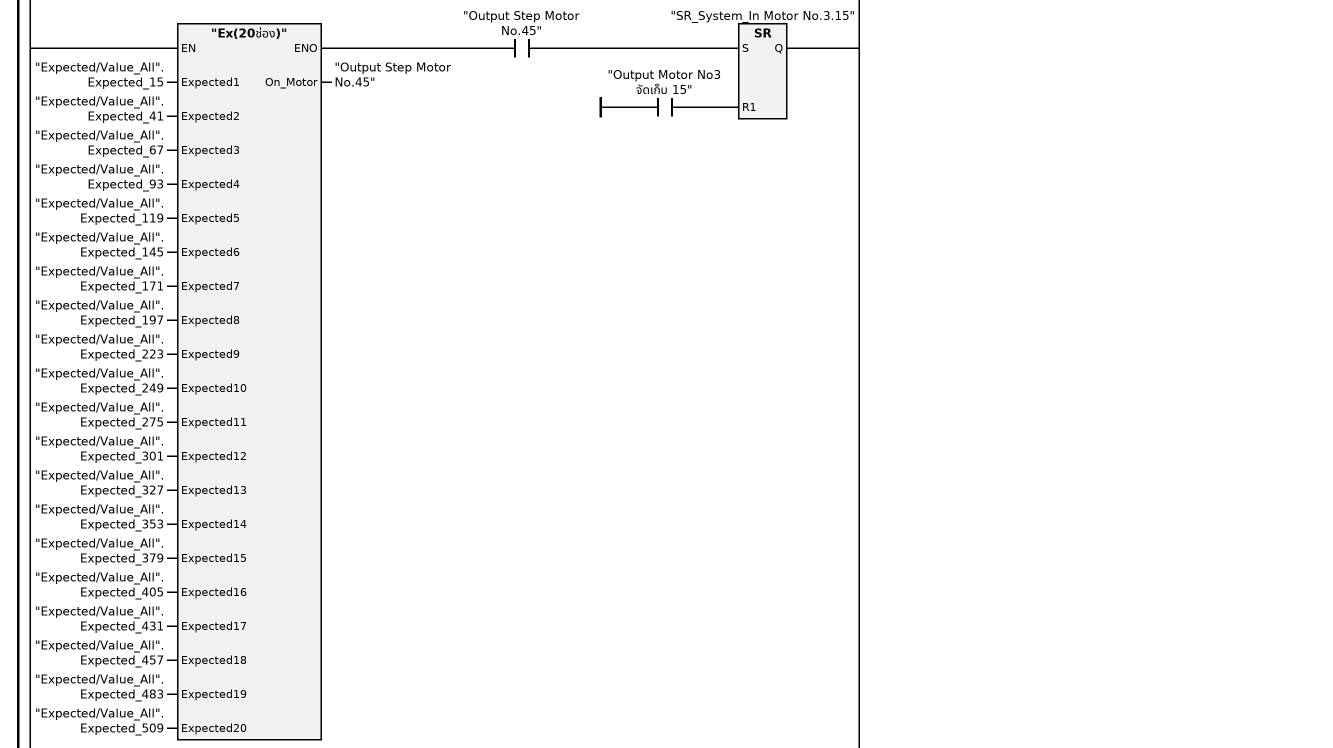
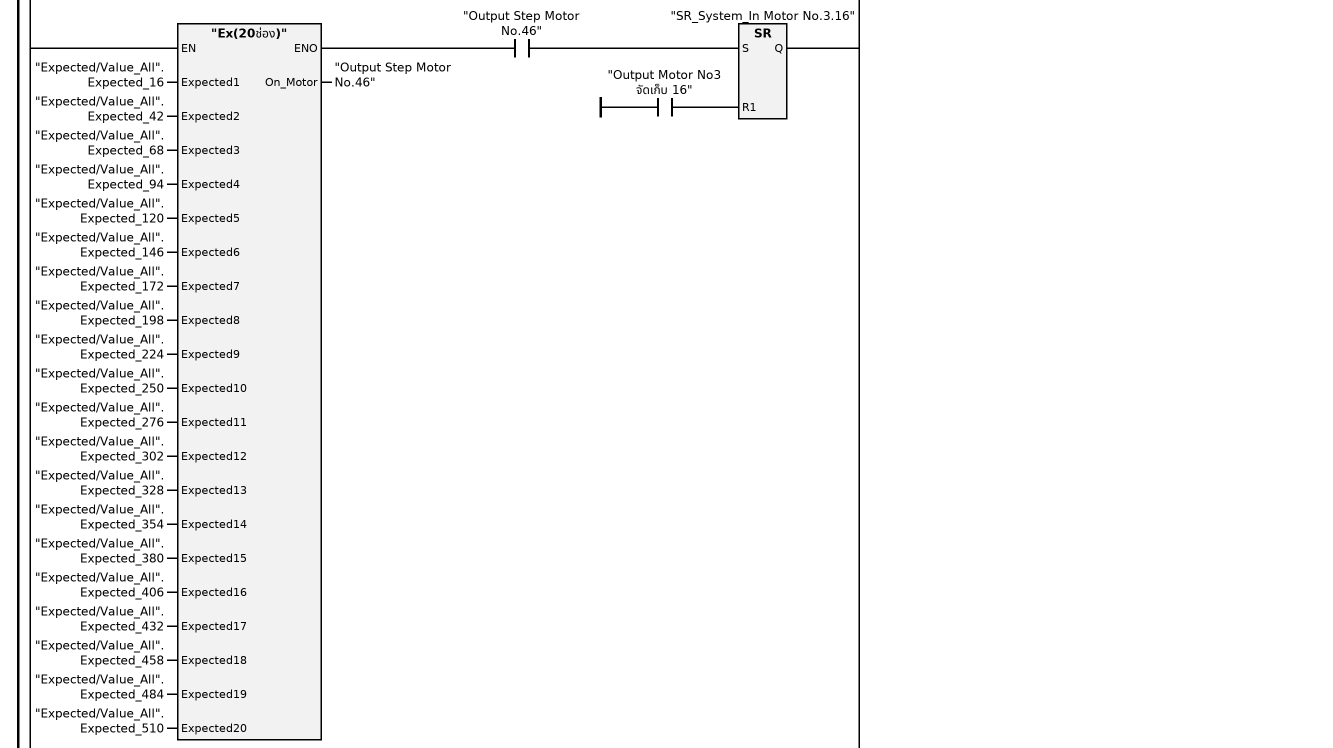
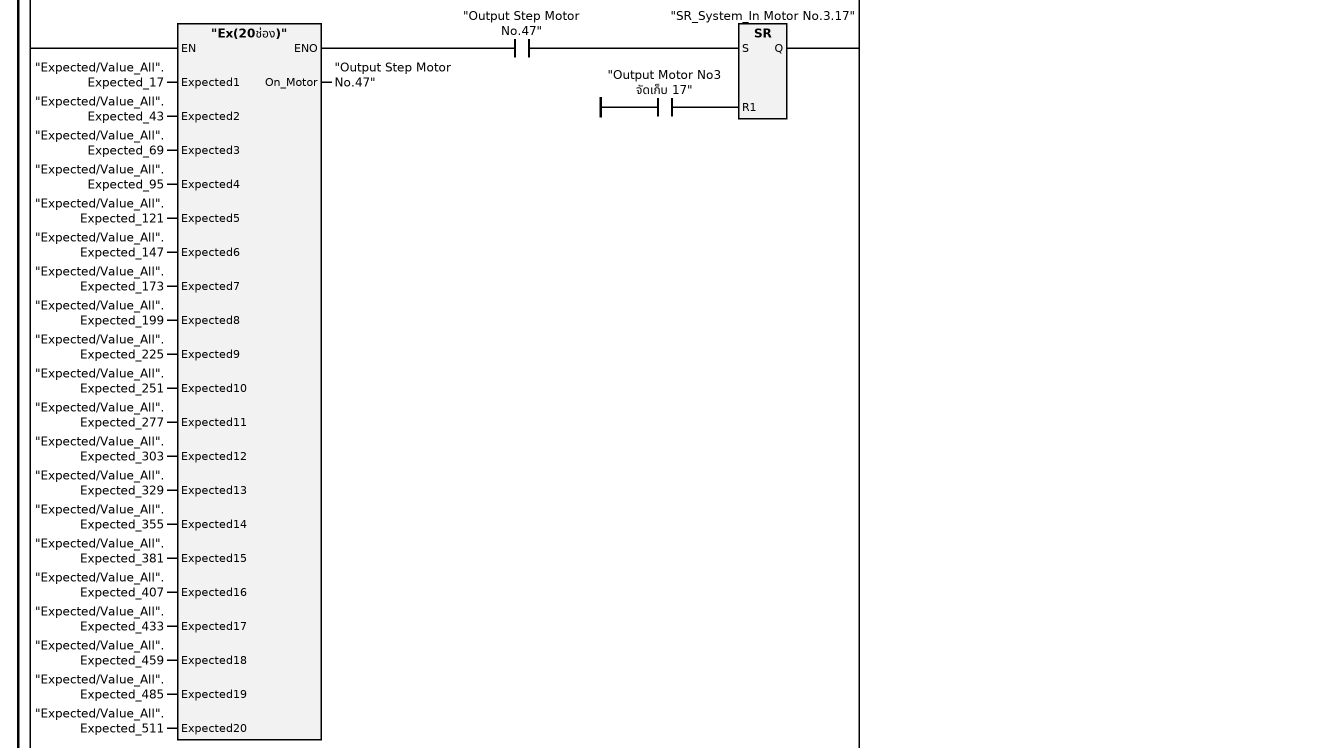
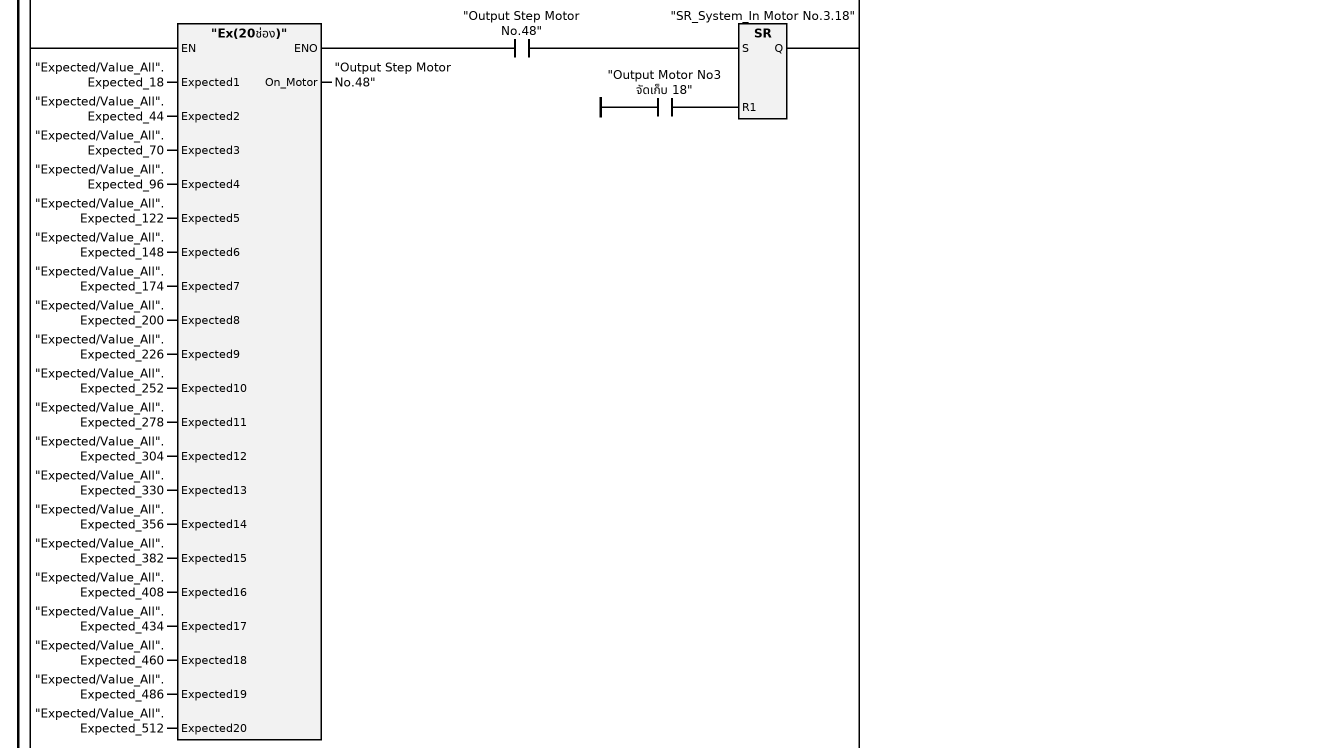
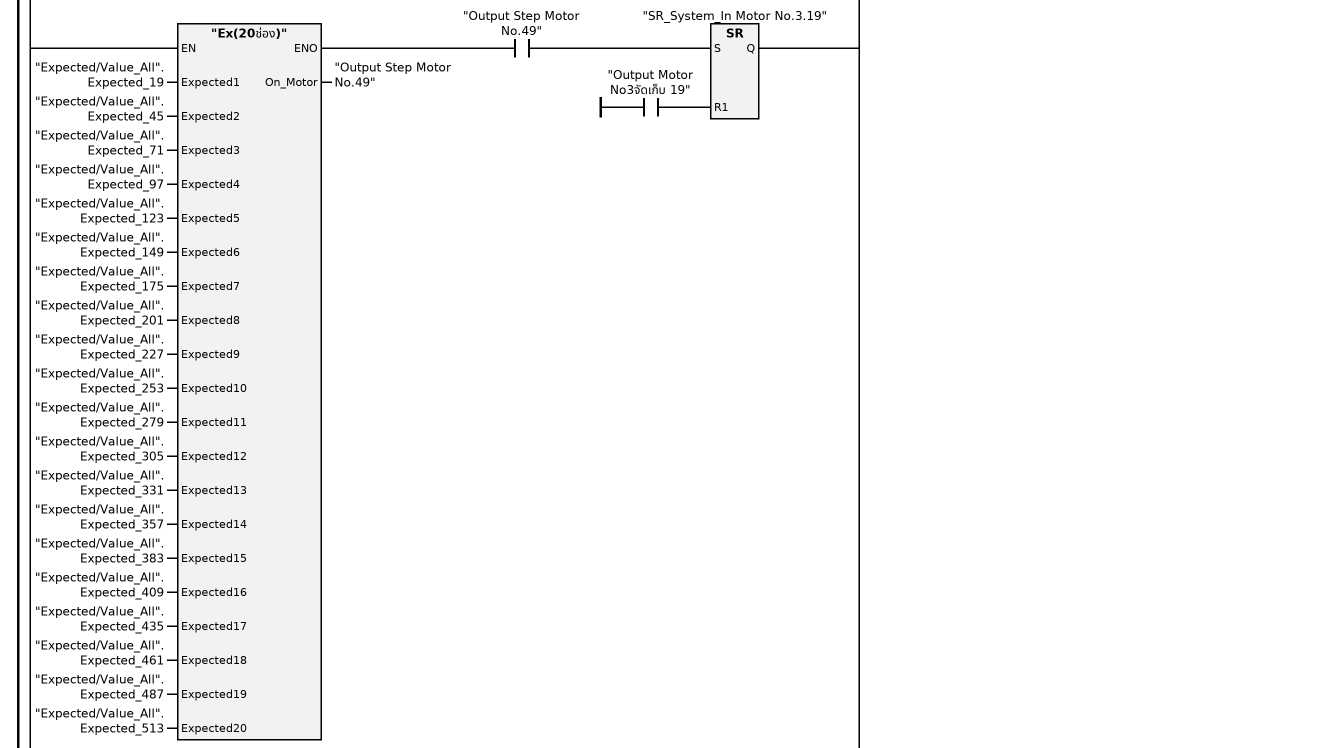
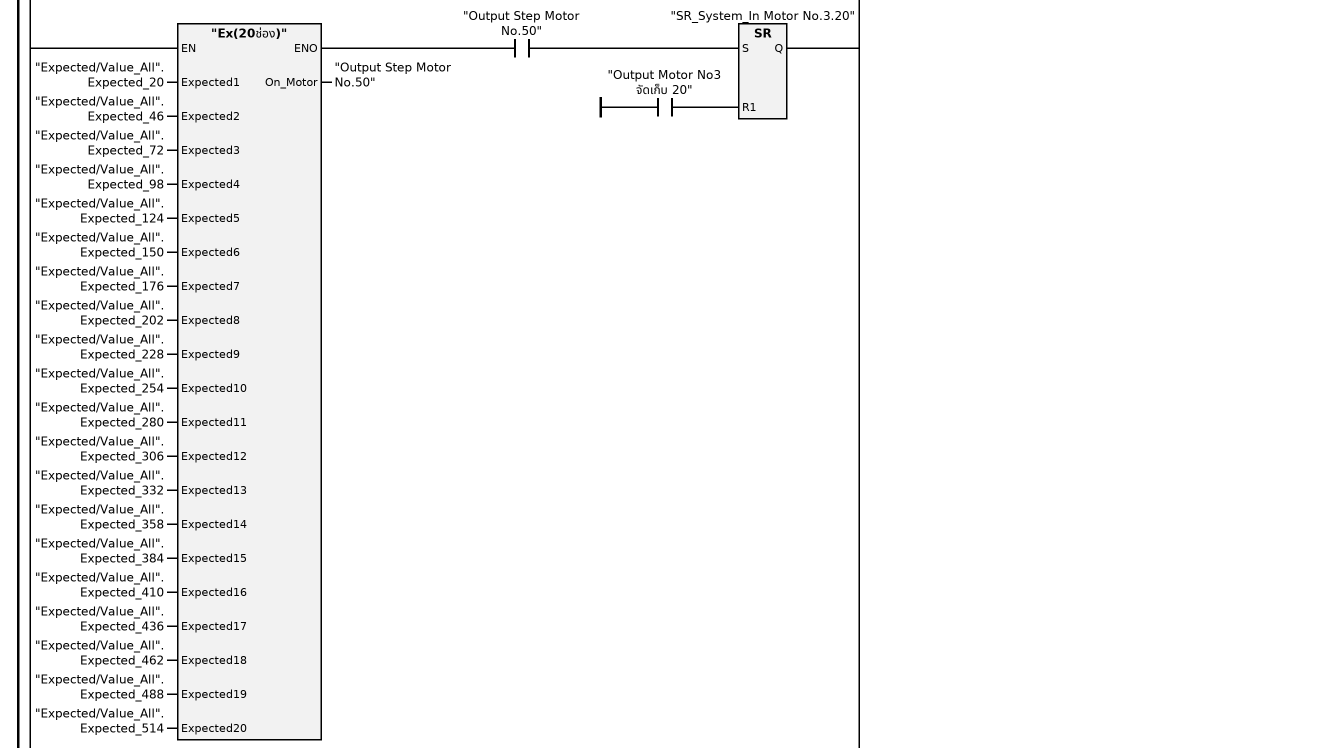
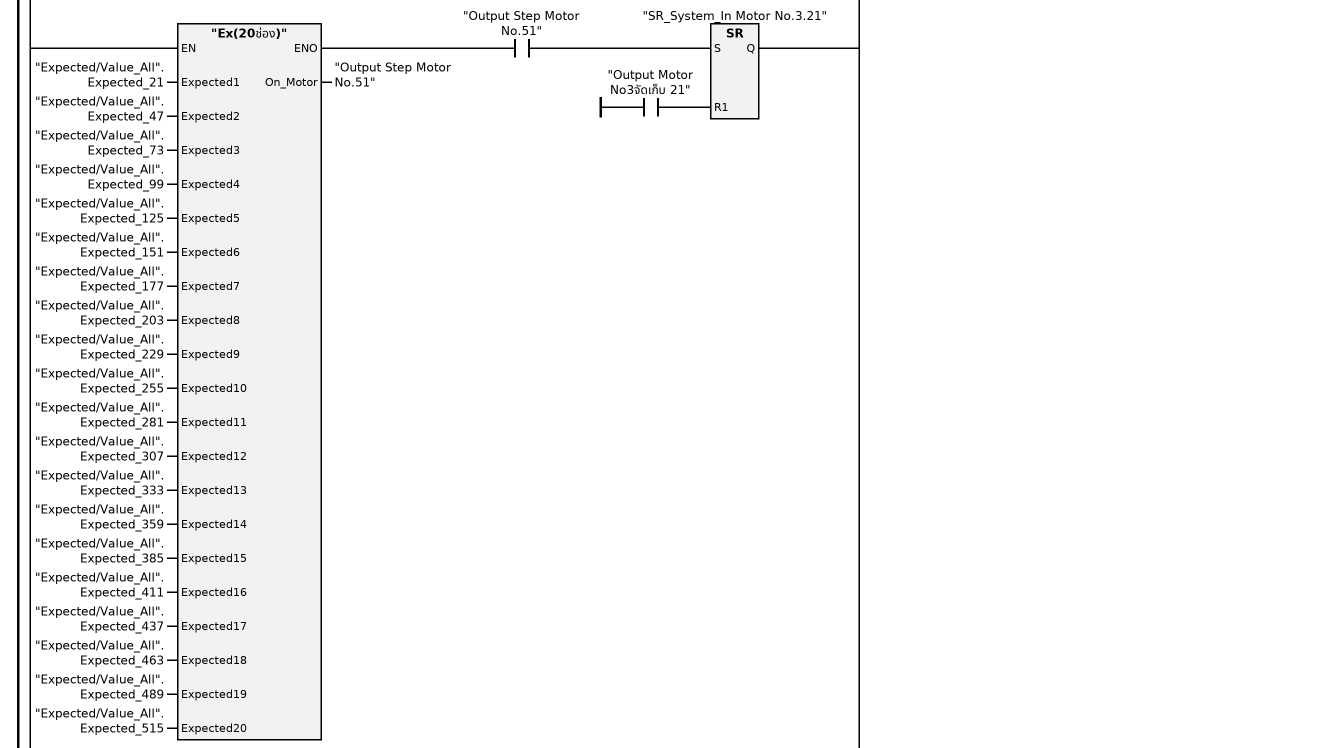
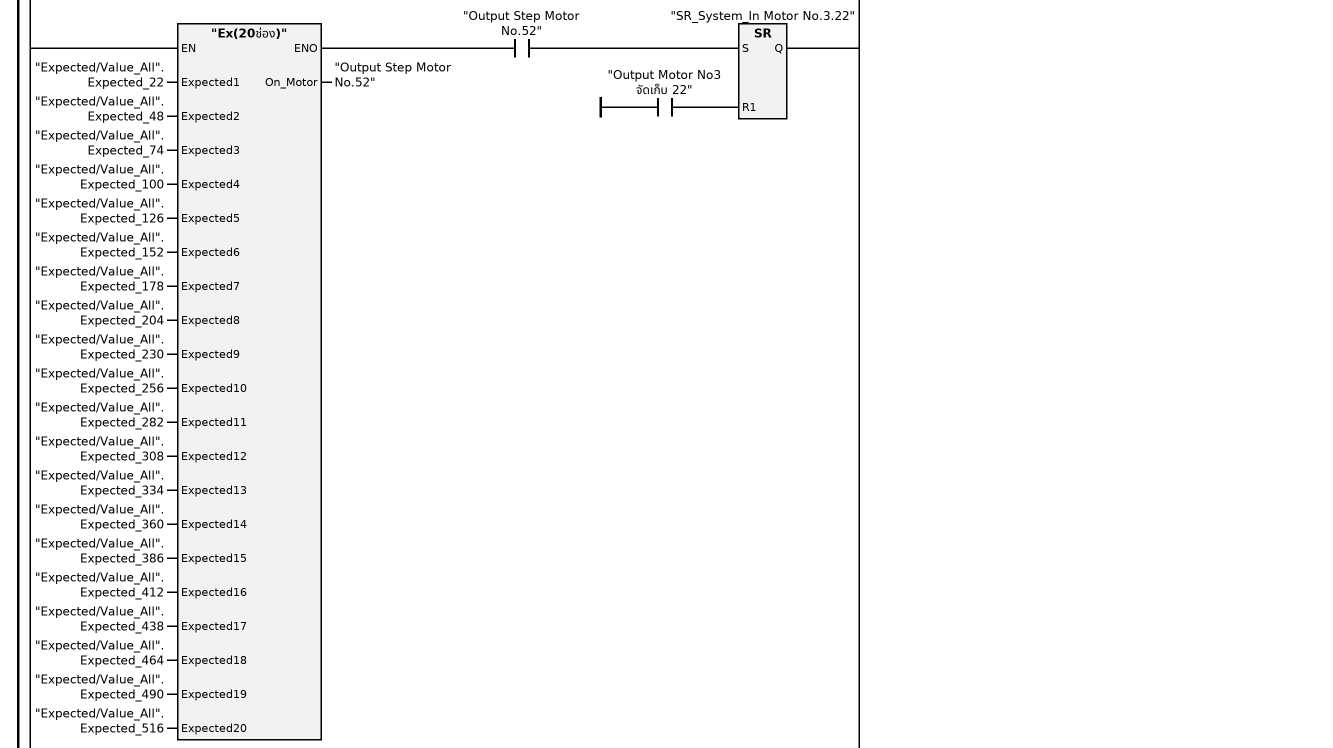
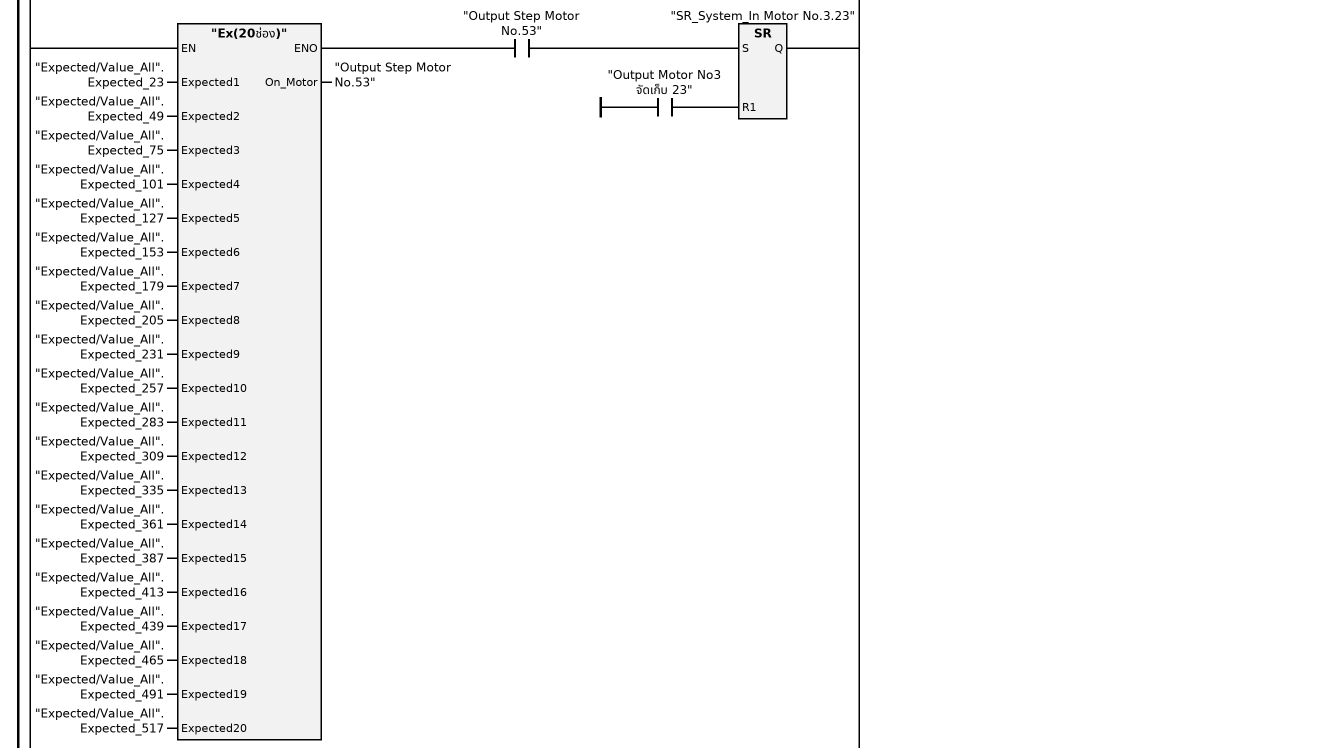
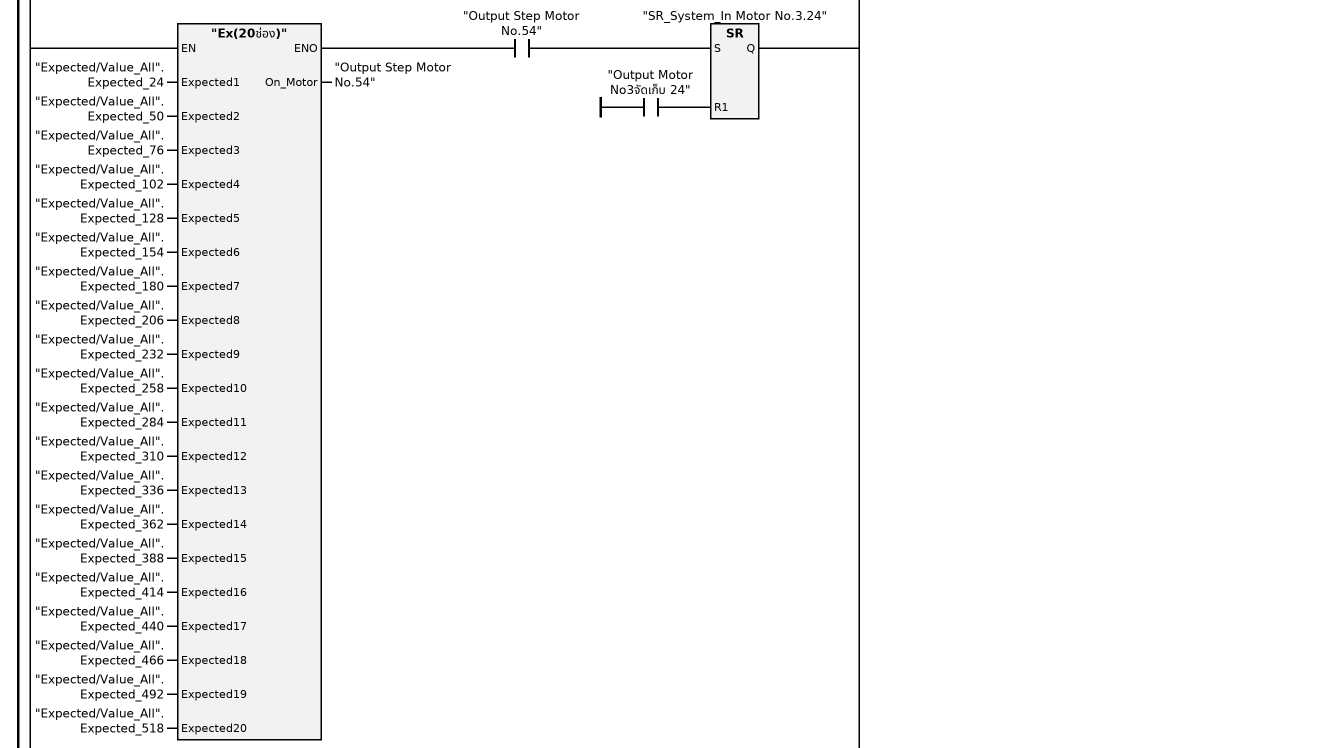
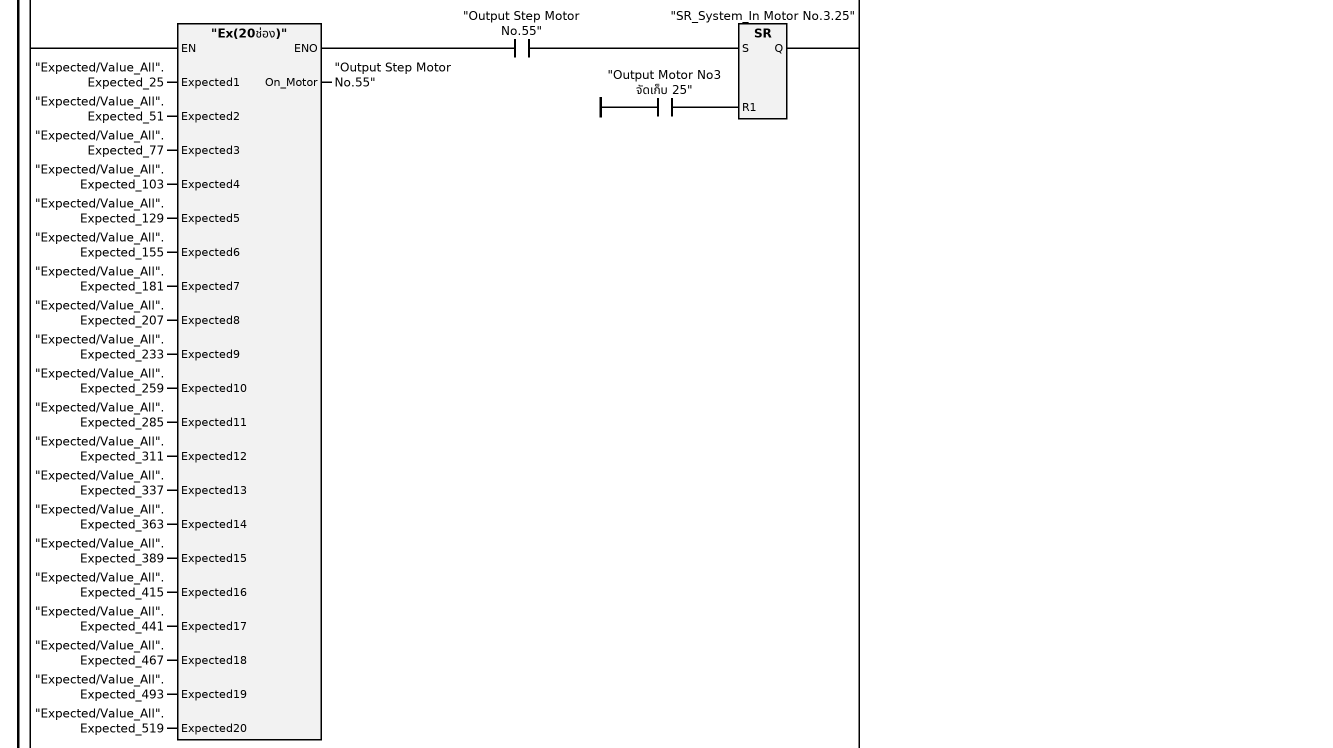
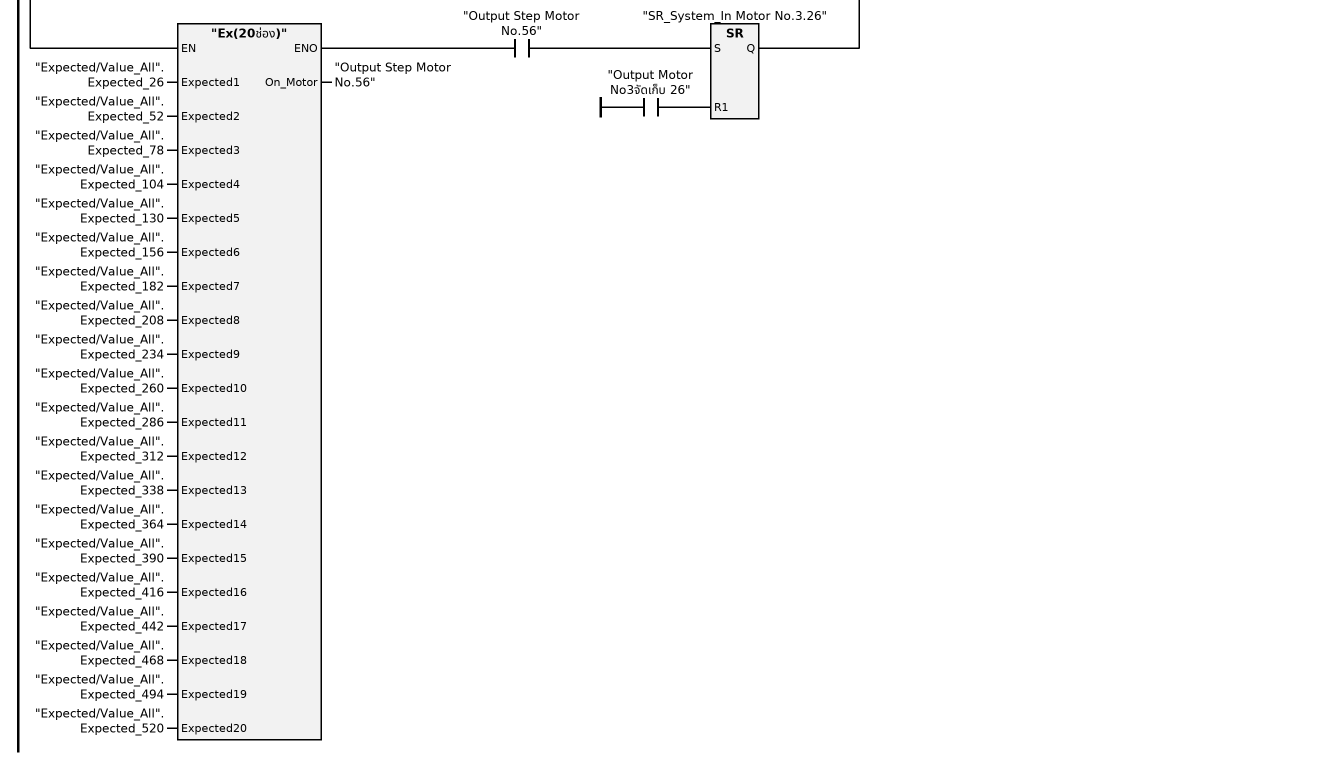
   "Ex(20ช่อง)"(Expected1 := "Expected/Value_All".Expected_1,
                Expected2 := "Expected/Value_All".Expected_27,
                Expected3 := "Expected/Value_All".Expected_53,
                Expected4 := "Expected/Value_All".Expected_79,
                Expected5 := "Expected/Value_All".Expected_105,
                Expected6 := "Expected/Value_All".Expected_131,
                Expected7 := "Expected/Value_All".Expected_157,
                Expected8 := "Expected/Value_All".Expected_183,
                Expected9 := "Expected/Value_All".Expected_209,
                Expected10 := "Expected/Value_All".Expected_235,
                Expected11 := "Expected/Value_All".Expected_261,
                Expected12 := "Expected/Value_All".Expected_287,
                Expected13 := "Expected/Value_All".Expected_313,
                Expected14 := "Expected/Value_All".Expected_339,
                Expected15 := "Expected/Value_All".Expected_365,
                Expected16 := "Expected/Value_All".Expected_391,
                Expected17 := "Expected/Value_All".Expected_417,
                Expected18 := "Expected/Value_All".Expected_443,
                Expected19 := "Expected/Value_All".Expected_469,
                Expected20 := "Expected/Value_All".Expected_495,
                On_Motor => "Output Step Motor No.31",
                ENO => #_w1);
   IF #_w1 AND "Output Step Motor No.31" THEN
       "SR_System_In Motor No.3.1" := TRUE;   // SR flip-flop
   END_IF;
   IF "Output Motor No3 จัดเก็บ 1" THEN "SR_System_In Motor No.3.1" := FALSE; END_IF;
   #_w3 := "SR_System_In Motor No.3.1";
   "Ex(20ช่อง)"(Expected1 := "Expected/Value_All".Expected_2,
                Expected2 := "Expected/Value_All".Expected_28,
                Expected3 := "Expected/Value_All".Expected_54,
                Expected4 := "Expected/Value_All".Expected_80,
                Expected5 := "Expected/Value_All".Expected_106,
                Expected6 := "Expected/Value_All".Expected_132,
                Expected7 := "Expected/Value_All".Expected_158,
                Expected8 := "Expected/Value_All".Expected_184,
                Expected9 := "Expected/Value_All".Expected_201,
                Expected10 := "Expected/Value_All".Expected_236,
                Expected11 := "Expected/Value_All".Expected_262,
                Expected12 := "Expected/Value_All".Expected_288,
                Expected13 := "Expected/Value_All".Expected_314,
                Expected14 := "Expected/Value_All".Expected_340,
                Expected15 := "Expected/Value_All".Expected_366,
                Expected16 := "Expected/Value_All".Expected_392,
                Expected17 := "Expected/Value_All".Expected_418,
                Expected18 := "Expected/Value_All".Expected_444,
                Expected19 := "Expected/Value_All".Expected_470,
                Expected20 := "Expected/Value_All".Expected_492,
                On_Motor => "Output Step Motor No.32",
                ENO => #_w2);
   IF #_w2 AND "Output Step Motor No.32" THEN
       "SR_System_In Motor No.3.2" := TRUE;   // SR flip-flop
   END_IF;
   IF "Output Motor No3 จัดเก็บ 2" THEN "SR_System_In Motor No.3.2" := FALSE; END_IF;
   #_w5 := "SR_System_In Motor No.3.2";
   "Ex(20ช่อง)"(Expected1 := "Expected/Value_All".Expected_3,
                Expected2 := "Expected/Value_All".Expected_29,
                Expected3 := "Expected/Value_All".Expected_55,
                Expected4 := "Expected/Value_All".Expected_81,
                Expected5 := "Expected/Value_All".Expected_107,
                Expected6 := "Expected/Value_All".Expected_133,
                Expected7 := "Expected/Value_All".Expected_159,
                Expected8 := "Expected/Value_All".Expected_185,
                Expected9 := "Expected/Value_All".Expected_211,
                Expected10 := "Expected/Value_All".Expected_237,
                Expected11 := "Expected/Value_All".Expected_263,
                Expected12 := "Expected/Value_All".Expected_289,
                Expected13 := "Expected/Value_All".Expected_315,
                Expected14 := "Expected/Value_All".Expected_341,
                Expected15 := "Expected/Value_All".Expected_367,
                Expected16 := "Expected/Value_All".Expected_393,
                Expected17 := "Expected/Value_All".Expected_419,
                Expected18 := "Expected/Value_All".Expected_445,
                Expected19 := "Expected/Value_All".Expected_471,
                Expected20 := "Expected/Value_All".Expected_497,
                On_Motor => "Output Step Motor No.33",
                ENO => #_w4);
   IF #_w4 AND "Output Step Motor No.33" THEN
       "SR_System_In Motor No.3.3" := TRUE;   // SR flip-flop
   END_IF;
   IF "Output Motor No3จัดเก็บ 3" THEN "SR_System_In Motor No.3.3" := FALSE; END_IF;
   #_w7 := "SR_System_In Motor No.3.3";
   "Ex(20ช่อง)"(Expected1 := "Expected/Value_All".Expected_4,
                Expected2 := "Expected/Value_All".Expected_30,
                Expected3 := "Expected/Value_All".Expected_56,
                Expected4 := "Expected/Value_All".Expected_82,
                Expected5 := "Expected/Value_All".Expected_108,
                Expected6 := "Expected/Value_All".Expected_134,
                Expected7 := "Expected/Value_All".Expected_160,
                Expected8 := "Expected/Value_All".Expected_186,
                Expected9 := "Expected/Value_All".Expected_212,
                Expected10 := "Expected/Value_All".Expected_238,
                Expected11 := "Expected/Value_All".Expected_264,
                Expected12 := "Expected/Value_All".Expected_290,
                Expected13 := "Expected/Value_All".Expected_316,
                Expected14 := "Expected/Value_All".Expected_342,
                Expected15 := "Expected/Value_All".Expected_368,
                Expected16 := "Expected/Value_All".Expected_394,
                Expected17 := "Expected/Value_All".Expected_420,
                Expected18 := "Expected/Value_All".Expected_446,
                Expected19 := "Expected/Value_All".Expected_472,
                Expected20 := "Expected/Value_All".Expected_498,
                On_Motor => "Output Step Motor No.34",
                ENO => #_w6);
   IF #_w6 AND "Output Step Motor No.34" THEN
       "SR_System_In Motor No.3.4" := TRUE;   // SR flip-flop
   END_IF;
   IF "Output Motor No3 จัดเก็บ 4" THEN "SR_System_In Motor No.3.4" := FALSE; END_IF;
   #_w9 := "SR_System_In Motor No.3.4";
   "Ex(20ช่อง)"(Expected1 := "Expected/Value_All".Expected_5,
                Expected2 := "Expected/Value_All".Expected_31,
                Expected3 := "Expected/Value_All".Expected_57,
                Expected4 := "Expected/Value_All".Expected_83,
                Expected5 := "Expected/Value_All".Expected_109,
                Expected6 := "Expected/Value_All".Expected_135,
                Expected7 := "Expected/Value_All".Expected_161,
                Expected8 := "Expected/Value_All".Expected_187,
                Expected9 := "Expected/Value_All".Expected_213,
                Expected10 := "Expected/Value_All".Expected_239,
                Expected11 := "Expected/Value_All".Expected_265,
                Expected12 := "Expected/Value_All".Expected_291,
                Expected13 := "Expected/Value_All".Expected_317,
                Expected14 := "Expected/Value_All".Expected_343,
                Expected15 := "Expected/Value_All".Expected_369,
                Expected16 := "Expected/Value_All".Expected_395,
                Expected17 := "Expected/Value_All".Expected_421,
                Expected18 := "Expected/Value_All".Expected_447,
                Expected19 := "Expected/Value_All".Expected_473,
                Expected20 := "Expected/Value_All".Expected_499,
                On_Motor => "Output Step Motor No.35",
                ENO => #_w8);
   IF #_w8 AND "Output Step Motor No.35" THEN
       "SR_System_In Motor No.3.5" := TRUE;   // SR flip-flop
   END_IF;
   IF "Output Motor No3จัดเก็บ 5" THEN "SR_System_In Motor No.3.5" := FALSE; END_IF;
   #_w11 := "SR_System_In Motor No.3.5";
   "Ex(20ช่อง)"(Expected1 := "Expected/Value_All".Expected_6,
                Expected2 := "Expected/Value_All".Expected_32,
                Expected3 := "Expected/Value_All".Expected_58,
                Expected4 := "Expected/Value_All".Expected_84,
                Expected5 := "Expected/Value_All".Expected_110,
                Expected6 := "Expected/Value_All".Expected_136,
                Expected7 := "Expected/Value_All".Expected_162,
                Expected8 := "Expected/Value_All".Expected_188,
                Expected9 := "Expected/Value_All".Expected_214,
                Expected10 := "Expected/Value_All".Expected_240,
                Expected11 := "Expected/Value_All".Expected_266,
                Expected12 := "Expected/Value_All".Expected_292,
                Expected13 := "Expected/Value_All".Expected_318,
                Expected14 := "Expected/Value_All".Expected_344,
                Expected15 := "Expected/Value_All".Expected_370,
                Expected16 := "Expected/Value_All".Expected_396,
                Expected17 := "Expected/Value_All".Expected_422,
                Expected18 := "Expected/Value_All".Expected_448,
                Expected19 := "Expected/Value_All".Expected_474,
                Expected20 := "Expected/Value_All".Expected_500,
                On_Motor => "Output Step Motor No.36",
                ENO => #_w10);
   IF #_w10 AND "Output Step Motor No.36" THEN
       "SR_System_In Motor No.3.6" := TRUE;   // SR flip-flop
   END_IF;
   IF "Output Motor No3 จัดเก็บ 6" THEN "SR_System_In Motor No.3.6" := FALSE; END_IF;
   #_w13 := "SR_System_In Motor No.3.6";
   "Ex(20ช่อง)"(Expected1 := "Expected/Value_All".Expected_7,
                Expected2 := "Expected/Value_All".Expected_33,
                Expected3 := "Expected/Value_All".Expected_59,
                Expected4 := "Expected/Value_All".Expected_85,
                Expected5 := "Expected/Value_All".Expected_111,
                Expected6 := "Expected/Value_All".Expected_137,
                Expected7 := "Expected/Value_All".Expected_163,
                Expected8 := "Expected/Value_All".Expected_189,
                Expected9 := "Expected/Value_All".Expected_215,
                Expected10 := "Expected/Value_All".Expected_241,
                Expected11 := "Expected/Value_All".Expected_267,
                Expected12 := "Expected/Value_All".Expected_293,
                Expected13 := "Expected/Value_All".Expected_319,
                Expected14 := "Expected/Value_All".Expected_345,
                Expected15 := "Expected/Value_All".Expected_371,
                Expected16 := "Expected/Value_All".Expected_397,
                Expected17 := "Expected/Value_All".Expected_423,
                Expected18 := "Expected/Value_All".Expected_449,
                Expected19 := "Expected/Value_All".Expected_475,
                Expected20 := "Expected/Value_All".Expected_501,
                On_Motor => "Output Step Motor No.37",
                ENO => #_w12);
   IF #_w12 AND "Output Step Motor No.37" THEN
       "SR_System_In Motor No.3.7" := TRUE;   // SR flip-flop
   END_IF;
   IF "Output Motor No3 จัดเก็บ 7" THEN "SR_System_In Motor No.3.7" := FALSE; END_IF;
   #_w15 := "SR_System_In Motor No.3.7";
   "Ex(20ช่อง)"(Expected1 := "Expected/Value_All".Expected_8,
                Expected2 := "Expected/Value_All".Expected_34,
                Expected3 := "Expected/Value_All".Expected_60,
                Expected4 := "Expected/Value_All".Expected_86,
                Expected5 := "Expected/Value_All".Expected_112,
                Expected6 := "Expected/Value_All".Expected_138,
                Expected7 := "Expected/Value_All".Expected_164,
                Expected8 := "Expected/Value_All".Expected_190,
                Expected9 := "Expected/Value_All".Expected_216,
                Expected10 := "Expected/Value_All".Expected_242,
                Expected11 := "Expected/Value_All".Expected_268,
                Expected12 := "Expected/Value_All".Expected_294,
                Expected13 := "Expected/Value_All".Expected_320,
                Expected14 := "Expected/Value_All".Expected_346,
                Expected15 := "Expected/Value_All".Expected_372,
                Expected16 := "Expected/Value_All".Expected_398,
                Expected17 := "Expected/Value_All".Expected_424,
                Expected18 := "Expected/Value_All".Expected_450,
                Expected19 := "Expected/Value_All".Expected_476,
                Expected20 := "Expected/Value_All".Expected_502,
                On_Motor => "Output Step Motor No.38",
                ENO => #_w14);
   IF #_w14 AND "Output Step Motor No.38" THEN
       "SR_System_In Motor No.3.8" := TRUE;   // SR flip-flop
   END_IF;
   IF "Output Motor No3 จัดเก็บ 8" THEN "SR_System_In Motor No.3.8" := FALSE; END_IF;
   #_w17 := "SR_System_In Motor No.3.8";
   "Ex(20ช่อง)"(Expected1 := "Expected/Value_All".Expected_9,
                Expected2 := "Expected/Value_All".Expected_35,
                Expected3 := "Expected/Value_All".Expected_61,
                Expected4 := "Expected/Value_All".Expected_87,
                Expected5 := "Expected/Value_All".Expected_113,
                Expected6 := "Expected/Value_All".Expected_139,
                Expected7 := "Expected/Value_All".Expected_165,
                Expected8 := "Expected/Value_All".Expected_191,
                Expected9 := "Expected/Value_All".Expected_217,
                Expected10 := "Expected/Value_All".Expected_243,
                Expected11 := "Expected/Value_All".Expected_269,
                Expected12 := "Expected/Value_All".Expected_295,
                Expected13 := "Expected/Value_All".Expected_321,
                Expected14 := "Expected/Value_All".Expected_347,
                Expected15 := "Expected/Value_All".Expected_373,
                Expected16 := "Expected/Value_All".Expected_399,
                Expected17 := "Expected/Value_All".Expected_425,
                Expected18 := "Expected/Value_All".Expected_451,
                Expected19 := "Expected/Value_All".Expected_477,
                Expected20 := "Expected/Value_All".Expected_503,
                On_Motor => "Output Step Motor No.39",
                ENO => #_w16);
   IF #_w16 AND "Output Step Motor No.39" THEN
       "SR_System_In Motor No.3.9" := TRUE;   // SR flip-flop
   END_IF;
   IF "Output Motor No3 จัดเก็บ 9" THEN "SR_System_In Motor No.3.9" := FALSE; END_IF;
   #_w19 := "SR_System_In Motor No.3.9";
   "Ex(20ช่อง)"(Expected1 := "Expected/Value_All".Expected_10,
                Expected2 := "Expected/Value_All".Expected_36,
                Expected3 := "Expected/Value_All".Expected_62,
                Expected4 := "Expected/Value_All".Expected_88,
                Expected5 := "Expected/Value_All".Expected_114,
                Expected6 := "Expected/Value_All".Expected_140,
                Expected7 := "Expected/Value_All".Expected_166,
                Expected8 := "Expected/Value_All".Expected_192,
                Expected9 := "Expected/Value_All".Expected_218,
                Expected10 := "Expected/Value_All".Expected_244,
                Expected11 := "Expected/Value_All".Expected_270,
                Expected12 := "Expected/Value_All".Expected_296,
                Expected13 := "Expected/Value_All".Expected_322,
                Expected14 := "Expected/Value_All".Expected_348,
                Expected15 := "Expected/Value_All".Expected_374,
                Expected16 := "Expected/Value_All".Expected_400,
                Expected17 := "Expected/Value_All".Expected_426,
                Expected18 := "Expected/Value_All".Expected_452,
                Expected19 := "Expected/Value_All".Expected_478,
                Expected20 := "Expected/Value_All".Expected_504,
                On_Motor => "Output Step Motor No.40",
                ENO => #_w18);
   IF #_w18 AND "Output Step Motor No.40" THEN
       "SR_System_In Motor No.3.10" := TRUE;   // SR flip-flop
   END_IF;
   IF "Output Motor No3 จัดเก็บ10" THEN "SR_System_In Motor No.3.10" := FALSE; END_IF;
   #_w21 := "SR_System_In Motor No.3.10";
   "Ex(20ช่อง)"(Expected1 := "Expected/Value_All".Expected_11,
                Expected2 := "Expected/Value_All".Expected_37,
                Expected3 := "Expected/Value_All".Expected_63,
                Expected4 := "Expected/Value_All".Expected_89,
                Expected5 := "Expected/Value_All".Expected_115,
                Expected6 := "Expected/Value_All".Expected_141,
                Expected7 := "Expected/Value_All".Expected_167,
                Expected8 := "Expected/Value_All".Expected_193,
                Expected9 := "Expected/Value_All".Expected_219,
                Expected10 := "Expected/Value_All".Expected_245,
                Expected11 := "Expected/Value_All".Expected_271,
                Expected12 := "Expected/Value_All".Expected_297,
                Expected13 := "Expected/Value_All".Expected_323,
                Expected14 := "Expected/Value_All".Expected_349,
                Expected15 := "Expected/Value_All".Expected_375,
                Expected16 := "Expected/Value_All".Expected_401,
                Expected17 := "Expected/Value_All".Expected_427,
                Expected18 := "Expected/Value_All".Expected_453,
                Expected19 := "Expected/Value_All".Expected_479,
                Expected20 := "Expected/Value_All".Expected_505,
                On_Motor => "Output Step Motor No.41",
                ENO => #_w20);
   IF #_w20 AND "Output Step Motor No.41" THEN
       "SR_System_In Motor No.3.11" := TRUE;   // SR flip-flop
   END_IF;
   IF "Output Motor No3จัดเก็บ 11" THEN "SR_System_In Motor No.3.11" := FALSE; END_IF;
   #_w23 := "SR_System_In Motor No.3.11";
   "Ex(20ช่อง)"(Expected1 := "Expected/Value_All".Expected_12,
                Expected2 := "Expected/Value_All".Expected_38,
                Expected3 := "Expected/Value_All".Expected_64,
                Expected4 := "Expected/Value_All".Expected_90,
                Expected5 := "Expected/Value_All".Expected_116,
                Expected6 := "Expected/Value_All".Expected_142,
                Expected7 := "Expected/Value_All".Expected_168,
                Expected8 := "Expected/Value_All".Expected_194,
                Expected9 := "Expected/Value_All".Expected_220,
                Expected10 := "Expected/Value_All".Expected_246,
                Expected11 := "Expected/Value_All".Expected_272,
                Expected12 := "Expected/Value_All".Expected_298,
                Expected13 := "Expected/Value_All".Expected_324,
                Expected14 := "Expected/Value_All".Expected_350,
                Expected15 := "Expected/Value_All".Expected_376,
                Expected16 := "Expected/Value_All".Expected_402,
                Expected17 := "Expected/Value_All".Expected_428,
                Expected18 := "Expected/Value_All".Expected_454,
                Expected19 := "Expected/Value_All".Expected_480,
                Expected20 := "Expected/Value_All".Expected_506,
                On_Motor => "Output Step Motor No.42",
                ENO => #_w22);
   IF #_w22 AND "Output Step Motor No.42" THEN
       "SR_System_In Motor No.3.12" := TRUE;   // SR flip-flop
   END_IF;
   IF "Output Motor No3 จัดเก็บ 12" THEN "SR_System_In Motor No.3.12" := FALSE; END_IF;
   #_w25 := "SR_System_In Motor No.3.12";
   "Ex(20ช่อง)"(Expected1 := "Expected/Value_All".Expected_13,
                Expected2 := "Expected/Value_All".Expected_39,
                Expected3 := "Expected/Value_All".Expected_65,
                Expected4 := "Expected/Value_All".Expected_91,
                Expected5 := "Expected/Value_All".Expected_117,
                Expected6 := "Expected/Value_All".Expected_143,
                Expected7 := "Expected/Value_All".Expected_169,
                Expected8 := "Expected/Value_All".Expected_195,
                Expected9 := "Expected/Value_All".Expected_221,
                Expected10 := "Expected/Value_All".Expected_247,
                Expected11 := "Expected/Value_All".Expected_273,
                Expected12 := "Expected/Value_All".Expected_299,
                Expected13 := "Expected/Value_All".Expected_325,
                Expected14 := "Expected/Value_All".Expected_351,
                Expected15 := "Expected/Value_All".Expected_377,
                Expected16 := "Expected/Value_All".Expected_403,
                Expected17 := "Expected/Value_All".Expected_429,
                Expected18 := "Expected/Value_All".Expected_455,
                Expected19 := "Expected/Value_All".Expected_481,
                Expected20 := "Expected/Value_All".Expected_507,
                On_Motor => "Output Step Motor No.43",
                ENO => #_w24);
   IF #_w24 AND "Output Step Motor No.43" THEN
       "SR_System_In Motor No.3.13" := TRUE;   // SR flip-flop
   END_IF;
   IF "Output Motor No3จัดเก็บ 13" THEN "SR_System_In Motor No.3.13" := FALSE; END_IF;
   #_w27 := "SR_System_In Motor No.3.13";
   "Ex(20ช่อง)"(Expected1 := "Expected/Value_All".Expected_14,
                Expected2 := "Expected/Value_All".Expected_40,
                Expected3 := "Expected/Value_All".Expected_66,
                Expected4 := "Expected/Value_All".Expected_92,
                Expected5 := "Expected/Value_All".Expected_118,
                Expected6 := "Expected/Value_All".Expected_144,
                Expected7 := "Expected/Value_All".Expected_170,
                Expected8 := "Expected/Value_All".Expected_196,
                Expected9 := "Expected/Value_All".Expected_222,
                Expected10 := "Expected/Value_All".Expected_248,
                Expected11 := "Expected/Value_All".Expected_274,
                Expected12 := "Expected/Value_All".Expected_300,
                Expected13 := "Expected/Value_All".Expected_326,
                Expected14 := "Expected/Value_All".Expected_352,
                Expected15 := "Expected/Value_All".Expected_378,
                Expected16 := "Expected/Value_All".Expected_404,
                Expected17 := "Expected/Value_All".Expected_430,
                Expected18 := "Expected/Value_All".Expected_456,
                Expected19 := "Expected/Value_All".Expected_482,
                Expected20 := "Expected/Value_All".Expected_508,
                On_Motor => "Output Step Motor No.44",
                ENO => #_w26);
   IF #_w26 AND "Output Step Motor No.44" THEN
       "SR_System_In Motor No.3.14" := TRUE;   // SR flip-flop
   END_IF;
   IF "Output Motor No3 จัดเก็บ 14" THEN "SR_System_In Motor No.3.14" := FALSE; END_IF;
   #_w29 := "SR_System_In Motor No.3.14";
   "Ex(20ช่อง)"(Expected1 := "Expected/Value_All".Expected_15,
                Expected2 := "Expected/Value_All".Expected_41,
                Expected3 := "Expected/Value_All".Expected_67,
                Expected4 := "Expected/Value_All".Expected_93,
                Expected5 := "Expected/Value_All".Expected_119,
                Expected6 := "Expected/Value_All".Expected_145,
                Expected7 := "Expected/Value_All".Expected_171,
                Expected8 := "Expected/Value_All".Expected_197,
                Expected9 := "Expected/Value_All".Expected_223,
                Expected10 := "Expected/Value_All".Expected_249,
                Expected11 := "Expected/Value_All".Expected_275,
                Expected12 := "Expected/Value_All".Expected_301,
                Expected13 := "Expected/Value_All".Expected_327,
                Expected14 := "Expected/Value_All".Expected_353,
                Expected15 := "Expected/Value_All".Expected_379,
                Expected16 := "Expected/Value_All".Expected_405,
                Expected17 := "Expected/Value_All".Expected_431,
                Expected18 := "Expected/Value_All".Expected_457,
                Expected19 := "Expected/Value_All".Expected_483,
                Expected20 := "Expected/Value_All".Expected_509,
                On_Motor => "Output Step Motor No.45",
                ENO => #_w28);
   IF #_w28 AND "Output Step Motor No.45" THEN
       "SR_System_In Motor No.3.15" := TRUE;   // SR flip-flop
   END_IF;
   IF "Output Motor No3 จัดเก็บ 15" THEN "SR_System_In Motor No.3.15" := FALSE; END_IF;
   #_w31 := "SR_System_In Motor No.3.15";
   "Ex(20ช่อง)"(Expected1 := "Expected/Value_All".Expected_16,
                Expected2 := "Expected/Value_All".Expected_42,
                Expected3 := "Expected/Value_All".Expected_68,
                Expected4 := "Expected/Value_All".Expected_94,
                Expected5 := "Expected/Value_All".Expected_120,
                Expected6 := "Expected/Value_All".Expected_146,
                Expected7 := "Expected/Value_All".Expected_172,
                Expected8 := "Expected/Value_All".Expected_198,
                Expected9 := "Expected/Value_All".Expected_224,
                Expected10 := "Expected/Value_All".Expected_250,
                Expected11 := "Expected/Value_All".Expected_276,
                Expected12 := "Expected/Value_All".Expected_302,
                Expected13 := "Expected/Value_All".Expected_328,
                Expected14 := "Expected/Value_All".Expected_354,
                Expected15 := "Expected/Value_All".Expected_380,
                Expected16 := "Expected/Value_All".Expected_406,
                Expected17 := "Expected/Value_All".Expected_432,
                Expected18 := "Expected/Value_All".Expected_458,
                Expected19 := "Expected/Value_All".Expected_484,
                Expected20 := "Expected/Value_All".Expected_510,
                On_Motor => "Output Step Motor No.46",
                ENO => #_w30);
   IF #_w30 AND "Output Step Motor No.46" THEN
       "SR_System_In Motor No.3.16" := TRUE;   // SR flip-flop
   END_IF;
   IF "Output Motor No3 จัดเก็บ 16" THEN "SR_System_In Motor No.3.16" := FALSE; END_IF;
   #_w33 := "SR_System_In Motor No.3.16";
   "Ex(20ช่อง)"(Expected1 := "Expected/Value_All".Expected_17,
                Expected2 := "Expected/Value_All".Expected_43,
                Expected3 := "Expected/Value_All".Expected_69,
                Expected4 := "Expected/Value_All".Expected_95,
                Expected5 := "Expected/Value_All".Expected_121,
                Expected6 := "Expected/Value_All".Expected_147,
                Expected7 := "Expected/Value_All".Expected_173,
                Expected8 := "Expected/Value_All".Expected_199,
                Expected9 := "Expected/Value_All".Expected_225,
                Expected10 := "Expected/Value_All".Expected_251,
                Expected11 := "Expected/Value_All".Expected_277,
                Expected12 := "Expected/Value_All".Expected_303,
                Expected13 := "Expected/Value_All".Expected_329,
                Expected14 := "Expected/Value_All".Expected_355,
                Expected15 := "Expected/Value_All".Expected_381,
                Expected16 := "Expected/Value_All".Expected_407,
                Expected17 := "Expected/Value_All".Expected_433,
                Expected18 := "Expected/Value_All".Expected_459,
                Expected19 := "Expected/Value_All".Expected_485,
                Expected20 := "Expected/Value_All".Expected_511,
                On_Motor => "Output Step Motor No.47",
                ENO => #_w32);
   IF #_w32 AND "Output Step Motor No.47" THEN
       "SR_System_In Motor No.3.17" := TRUE;   // SR flip-flop
   END_IF;
   IF "Output Motor No3 จัดเก็บ 17" THEN "SR_System_In Motor No.3.17" := FALSE; END_IF;
   #_w35 := "SR_System_In Motor No.3.17";
   "Ex(20ช่อง)"(Expected1 := "Expected/Value_All".Expected_18,
                Expected2 := "Expected/Value_All".Expected_44,
                Expected3 := "Expected/Value_All".Expected_70,
                Expected4 := "Expected/Value_All".Expected_96,
                Expected5 := "Expected/Value_All".Expected_122,
                Expected6 := "Expected/Value_All".Expected_148,
                Expected7 := "Expected/Value_All".Expected_174,
                Expected8 := "Expected/Value_All".Expected_200,
                Expected9 := "Expected/Value_All".Expected_226,
                Expected10 := "Expected/Value_All".Expected_252,
                Expected11 := "Expected/Value_All".Expected_278,
                Expected12 := "Expected/Value_All".Expected_304,
                Expected13 := "Expected/Value_All".Expected_330,
                Expected14 := "Expected/Value_All".Expected_356,
                Expected15 := "Expected/Value_All".Expected_382,
                Expected16 := "Expected/Value_All".Expected_408,
                Expected17 := "Expected/Value_All".Expected_434,
                Expected18 := "Expected/Value_All".Expected_460,
                Expected19 := "Expected/Value_All".Expected_486,
                Expected20 := "Expected/Value_All".Expected_512,
                On_Motor => "Output Step Motor No.48",
                ENO => #_w34);
   IF #_w34 AND "Output Step Motor No.48" THEN
       "SR_System_In Motor No.3.18" := TRUE;   // SR flip-flop
   END_IF;
   IF "Output Motor No3 จัดเก็บ 18" THEN "SR_System_In Motor No.3.18" := FALSE; END_IF;
   #_w37 := "SR_System_In Motor No.3.18";
   "Ex(20ช่อง)"(Expected1 := "Expected/Value_All".Expected_19,
                Expected2 := "Expected/Value_All".Expected_45,
                Expected3 := "Expected/Value_All".Expected_71,
                Expected4 := "Expected/Value_All".Expected_97,
                Expected5 := "Expected/Value_All".Expected_123,
                Expected6 := "Expected/Value_All".Expected_149,
                Expected7 := "Expected/Value_All".Expected_175,
                Expected8 := "Expected/Value_All".Expected_201,
                Expected9 := "Expected/Value_All".Expected_227,
                Expected10 := "Expected/Value_All".Expected_253,
                Expected11 := "Expected/Value_All".Expected_279,
                Expected12 := "Expected/Value_All".Expected_305,
                Expected13 := "Expected/Value_All".Expected_331,
                Expected14 := "Expected/Value_All".Expected_357,
                Expected15 := "Expected/Value_All".Expected_383,
                Expected16 := "Expected/Value_All".Expected_409,
                Expected17 := "Expected/Value_All".Expected_435,
                Expected18 := "Expected/Value_All".Expected_461,
                Expected19 := "Expected/Value_All".Expected_487,
                Expected20 := "Expected/Value_All".Expected_513,
                On_Motor => "Output Step Motor No.49",
                ENO => #_w36);
   IF #_w36 AND "Output Step Motor No.49" THEN
       "SR_System_In Motor No.3.19" := TRUE;   // SR flip-flop
   END_IF;
   IF "Output Motor No3จัดเก็บ 19" THEN "SR_System_In Motor No.3.19" := FALSE; END_IF;
   #_w39 := "SR_System_In Motor No.3.19";
   "Ex(20ช่อง)"(Expected1 := "Expected/Value_All".Expected_20,
                Expected2 := "Expected/Value_All".Expected_46,
                Expected3 := "Expected/Value_All".Expected_72,
                Expected4 := "Expected/Value_All".Expected_98,
                Expected5 := "Expected/Value_All".Expected_124,
                Expected6 := "Expected/Value_All".Expected_150,
                Expected7 := "Expected/Value_All".Expected_176,
                Expected8 := "Expected/Value_All".Expected_202,
                Expected9 := "Expected/Value_All".Expected_228,
                Expected10 := "Expected/Value_All".Expected_254,
                Expected11 := "Expected/Value_All".Expected_280,
                Expected12 := "Expected/Value_All".Expected_306,
                Expected13 := "Expected/Value_All".Expected_332,
                Expected14 := "Expected/Value_All".Expected_358,
                Expected15 := "Expected/Value_All".Expected_384,
                Expected16 := "Expected/Value_All".Expected_410,
                Expected17 := "Expected/Value_All".Expected_436,
                Expected18 := "Expected/Value_All".Expected_462,
                Expected19 := "Expected/Value_All".Expected_488,
                Expected20 := "Expected/Value_All".Expected_514,
                On_Motor => "Output Step Motor No.50",
                ENO => #_w38);
   IF #_w38 AND "Output Step Motor No.50" THEN
       "SR_System_In Motor No.3.20" := TRUE;   // SR flip-flop
   END_IF;
   IF "Output Motor No3 จัดเก็บ 20" THEN "SR_System_In Motor No.3.20" := FALSE; END_IF;
   #_w41 := "SR_System_In Motor No.3.20";
   "Ex(20ช่อง)"(Expected1 := "Expected/Value_All".Expected_21,
                Expected2 := "Expected/Value_All".Expected_47,
                Expected3 := "Expected/Value_All".Expected_73,
                Expected4 := "Expected/Value_All".Expected_99,
                Expected5 := "Expected/Value_All".Expected_125,
                Expected6 := "Expected/Value_All".Expected_151,
                Expected7 := "Expected/Value_All".Expected_177,
                Expected8 := "Expected/Value_All".Expected_203,
                Expected9 := "Expected/Value_All".Expected_229,
                Expected10 := "Expected/Value_All".Expected_255,
                Expected11 := "Expected/Value_All".Expected_281,
                Expected12 := "Expected/Value_All".Expected_307,
                Expected13 := "Expected/Value_All".Expected_333,
                Expected14 := "Expected/Value_All".Expected_359,
                Expected15 := "Expected/Value_All".Expected_385,
                Expected16 := "Expected/Value_All".Expected_411,
                Expected17 := "Expected/Value_All".Expected_437,
                Expected18 := "Expected/Value_All".Expected_463,
                Expected19 := "Expected/Value_All".Expected_489,
                Expected20 := "Expected/Value_All".Expected_515,
                On_Motor => "Output Step Motor No.51",
                ENO => #_w40);
   IF #_w40 AND "Output Step Motor No.51" THEN
       "SR_System_In Motor No.3.21" := TRUE;   // SR flip-flop
   END_IF;
   IF "Output Motor No3จัดเก็บ 21" THEN "SR_System_In Motor No.3.21" := FALSE; END_IF;
   #_w43 := "SR_System_In Motor No.3.21";
   "Ex(20ช่อง)"(Expected1 := "Expected/Value_All".Expected_22,
                Expected2 := "Expected/Value_All".Expected_48,
                Expected3 := "Expected/Value_All".Expected_74,
                Expected4 := "Expected/Value_All".Expected_100,
                Expected5 := "Expected/Value_All".Expected_126,
                Expected6 := "Expected/Value_All".Expected_152,
                Expected7 := "Expected/Value_All".Expected_178,
                Expected8 := "Expected/Value_All".Expected_204,
                Expected9 := "Expected/Value_All".Expected_230,
                Expected10 := "Expected/Value_All".Expected_256,
                Expected11 := "Expected/Value_All".Expected_282,
                Expected12 := "Expected/Value_All".Expected_308,
                Expected13 := "Expected/Value_All".Expected_334,
                Expected14 := "Expected/Value_All".Expected_360,
                Expected15 := "Expected/Value_All".Expected_386,
                Expected16 := "Expected/Value_All".Expected_412,
                Expected17 := "Expected/Value_All".Expected_438,
                Expected18 := "Expected/Value_All".Expected_464,
                Expected19 := "Expected/Value_All".Expected_490,
                Expected20 := "Expected/Value_All".Expected_516,
                On_Motor => "Output Step Motor No.52",
                ENO => #_w42);
   IF #_w42 AND "Output Step Motor No.52" THEN
       "SR_System_In Motor No.3.22" := TRUE;   // SR flip-flop
   END_IF;
   IF "Output Motor No3 จัดเก็บ 22" THEN "SR_System_In Motor No.3.22" := FALSE; END_IF;
   #_w45 := "SR_System_In Motor No.3.22";
   "Ex(20ช่อง)"(Expected1 := "Expected/Value_All".Expected_23,
                Expected2 := "Expected/Value_All".Expected_49,
                Expected3 := "Expected/Value_All".Expected_75,
                Expected4 := "Expected/Value_All".Expected_101,
                Expected5 := "Expected/Value_All".Expected_127,
                Expected6 := "Expected/Value_All".Expected_153,
                Expected7 := "Expected/Value_All".Expected_179,
                Expected8 := "Expected/Value_All".Expected_205,
                Expected9 := "Expected/Value_All".Expected_231,
                Expected10 := "Expected/Value_All".Expected_257,
                Expected11 := "Expected/Value_All".Expected_283,
                Expected12 := "Expected/Value_All".Expected_309,
                Expected13 := "Expected/Value_All".Expected_335,
                Expected14 := "Expected/Value_All".Expected_361,
                Expected15 := "Expected/Value_All".Expected_387,
                Expected16 := "Expected/Value_All".Expected_413,
                Expected17 := "Expected/Value_All".Expected_439,
                Expected18 := "Expected/Value_All".Expected_465,
                Expected19 := "Expected/Value_All".Expected_491,
                Expected20 := "Expected/Value_All".Expected_517,
                On_Motor => "Output Step Motor No.53",
                ENO => #_w44);
   IF #_w44 AND "Output Step Motor No.53" THEN
       "SR_System_In Motor No.3.23" := TRUE;   // SR flip-flop
   END_IF;
   IF "Output Motor No3 จัดเก็บ 23" THEN "SR_System_In Motor No.3.23" := FALSE; END_IF;
   #_w47 := "SR_System_In Motor No.3.23";
   "Ex(20ช่อง)"(Expected1 := "Expected/Value_All".Expected_24,
                Expected2 := "Expected/Value_All".Expected_50,
                Expected3 := "Expected/Value_All".Expected_76,
                Expected4 := "Expected/Value_All".Expected_102,
                Expected5 := "Expected/Value_All".Expected_128,
                Expected6 := "Expected/Value_All".Expected_154,
                Expected7 := "Expected/Value_All".Expected_180,
                Expected8 := "Expected/Value_All".Expected_206,
                Expected9 := "Expected/Value_All".Expected_232,
                Expected10 := "Expected/Value_All".Expected_258,
                Expected11 := "Expected/Value_All".Expected_284,
                Expected12 := "Expected/Value_All".Expected_310,
                Expected13 := "Expected/Value_All".Expected_336,
                Expected14 := "Expected/Value_All".Expected_362,
                Expected15 := "Expected/Value_All".Expected_388,
                Expected16 := "Expected/Value_All".Expected_414,
                Expected17 := "Expected/Value_All".Expected_440,
                Expected18 := "Expected/Value_All".Expected_466,
                Expected19 := "Expected/Value_All".Expected_492,
                Expected20 := "Expected/Value_All".Expected_518,
                On_Motor => "Output Step Motor No.54",
                ENO => #_w46);
   IF #_w46 AND "Output Step Motor No.54" THEN
       "SR_System_In Motor No.3.24" := TRUE;   // SR flip-flop
   END_IF;
   IF "Output Motor No3จัดเก็บ 24" THEN "SR_System_In Motor No.3.24" := FALSE; END_IF;
   #_w49 := "SR_System_In Motor No.3.24";
   "Ex(20ช่อง)"(Expected1 := "Expected/Value_All".Expected_25,
                Expected2 := "Expected/Value_All".Expected_51,
                Expected3 := "Expected/Value_All".Expected_77,
                Expected4 := "Expected/Value_All".Expected_103,
                Expected5 := "Expected/Value_All".Expected_129,
                Expected6 := "Expected/Value_All".Expected_155,
                Expected7 := "Expected/Value_All".Expected_181,
                Expected8 := "Expected/Value_All".Expected_207,
                Expected9 := "Expected/Value_All".Expected_233,
                Expected10 := "Expected/Value_All".Expected_259,
                Expected11 := "Expected/Value_All".Expected_285,
                Expected12 := "Expected/Value_All".Expected_311,
                Expected13 := "Expected/Value_All".Expected_337,
                Expected14 := "Expected/Value_All".Expected_363,
                Expected15 := "Expected/Value_All".Expected_389,
                Expected16 := "Expected/Value_All".Expected_415,
                Expected17 := "Expected/Value_All".Expected_441,
                Expected18 := "Expected/Value_All".Expected_467,
                Expected19 := "Expected/Value_All".Expected_493,
                Expected20 := "Expected/Value_All".Expected_519,
                On_Motor => "Output Step Motor No.55",
                ENO => #_w48);
   IF #_w48 AND "Output Step Motor No.55" THEN
       "SR_System_In Motor No.3.25" := TRUE;   // SR flip-flop
   END_IF;
   IF "Output Motor No3 จัดเก็บ 25" THEN "SR_System_In Motor No.3.25" := FALSE; END_IF;
   #_w51 := "SR_System_In Motor No.3.25";
   "Ex(20ช่อง)"(Expected1 := "Expected/Value_All".Expected_26,
                Expected2 := "Expected/Value_All".Expected_52,
                Expected3 := "Expected/Value_All".Expected_78,
                Expected4 := "Expected/Value_All".Expected_104,
                Expected5 := "Expected/Value_All".Expected_130,
                Expected6 := "Expected/Value_All".Expected_156,
                Expected7 := "Expected/Value_All".Expected_182,
                Expected8 := "Expected/Value_All".Expected_208,
                Expected9 := "Expected/Value_All".Expected_234,
                Expected10 := "Expected/Value_All".Expected_260,
                Expected11 := "Expected/Value_All".Expected_286,
                Expected12 := "Expected/Value_All".Expected_312,
                Expected13 := "Expected/Value_All".Expected_338,
                Expected14 := "Expected/Value_All".Expected_364,
                Expected15 := "Expected/Value_All".Expected_390,
                Expected16 := "Expected/Value_All".Expected_416,
                Expected17 := "Expected/Value_All".Expected_442,
                Expected18 := "Expected/Value_All".Expected_468,
                Expected19 := "Expected/Value_All".Expected_494,
                Expected20 := "Expected/Value_All".Expected_520,
                On_Motor => "Output Step Motor No.56",
                ENO => #_w50);
   IF #_w50 AND "Output Step Motor No.56" THEN
       "SR_System_In Motor No.3.26" := TRUE;   // SR flip-flop
   END_IF;
   IF "Output Motor No3จัดเก็บ 26" THEN "SR_System_In Motor No.3.26" := FALSE; END_IF;
   "IEC_Counter_0_DB_1593".CTU(CU := (#_w3 OR #_w5 OR #_w7 OR #_w9 OR #_w11 OR #_w13 OR #_w15 OR #_w17 OR #_w19 OR #_w21 OR #_w23 OR #_w25 OR #_w27 OR #_w29 OR #_w31 OR #_w33 OR #_w35 OR #_w37 OR #_w39 OR #_w41 OR #_w43 OR #_w45 OR #_w47 OR #_w49 OR #_w51 OR "SR_System_In Motor No.3.26") AND "Output test1",
                           R := "Outputtest2",
                           PV := 1);
   #"Stepper Motor  ทำงาน3" := "IEC_Counter_0_DB_1593".Q;
END_REGION

REGION Network 2
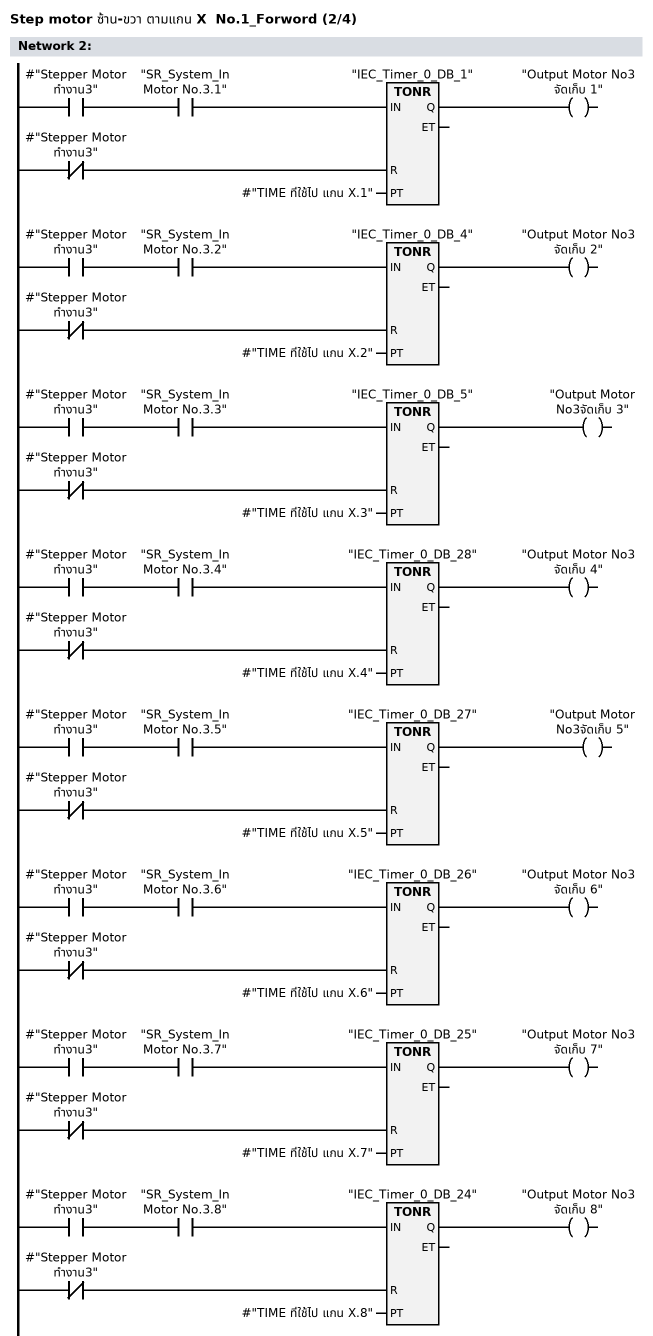
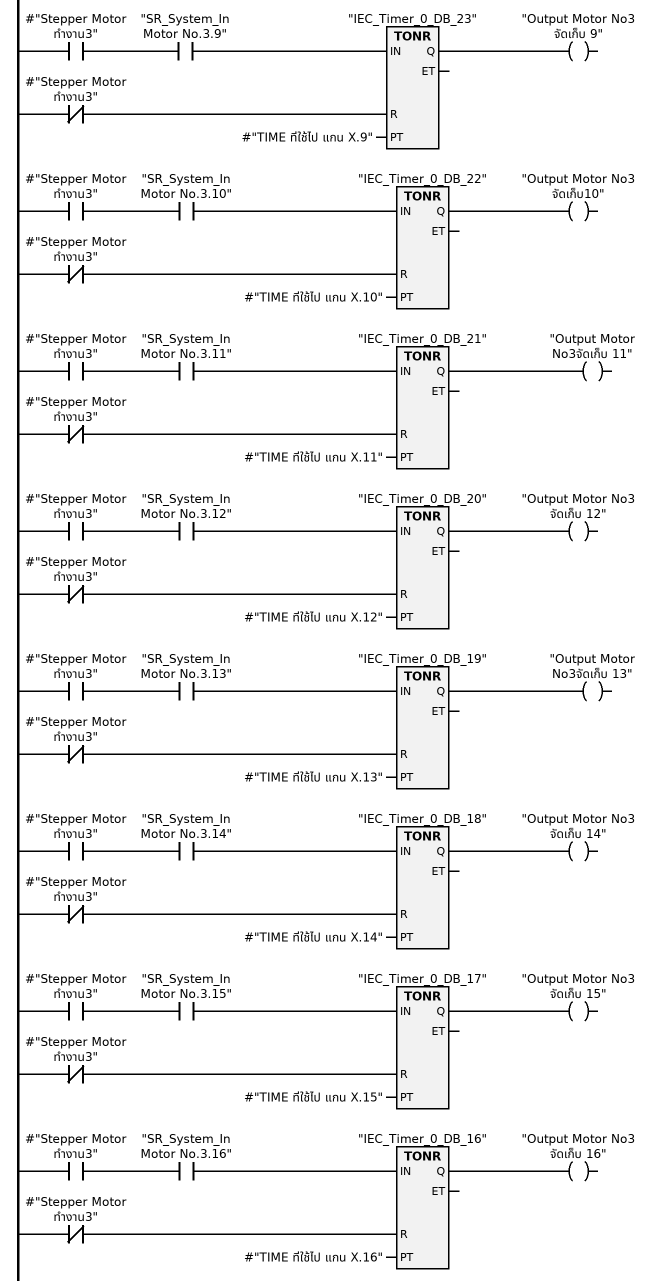
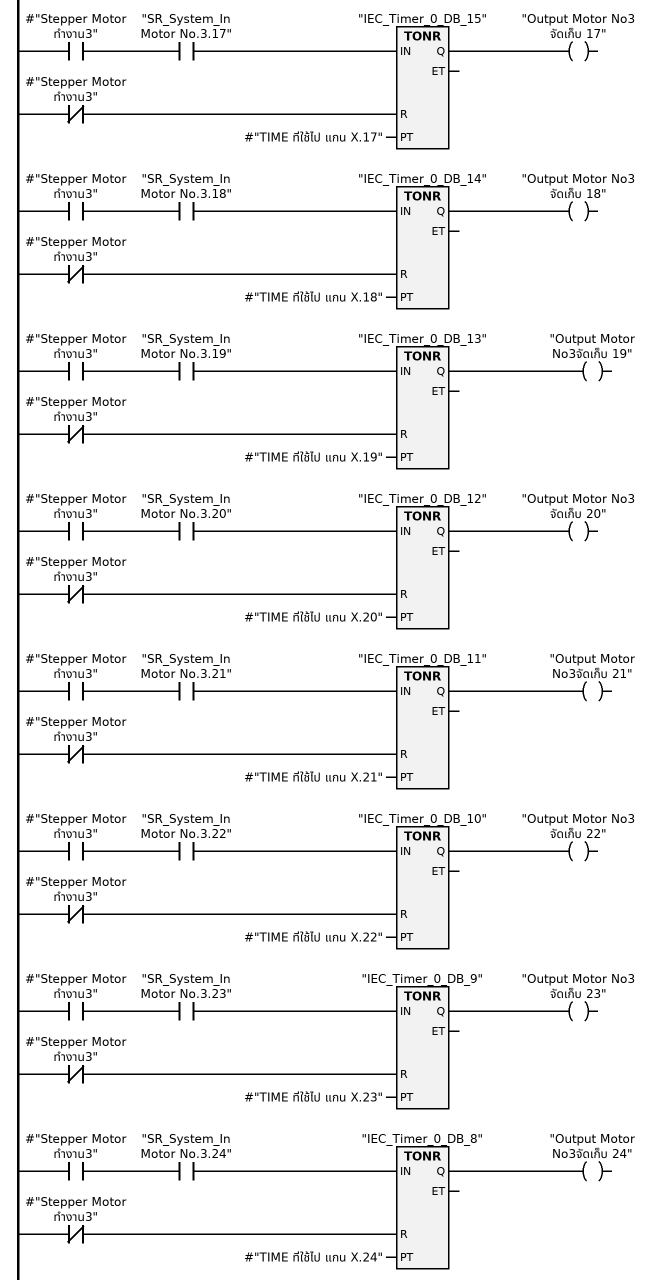
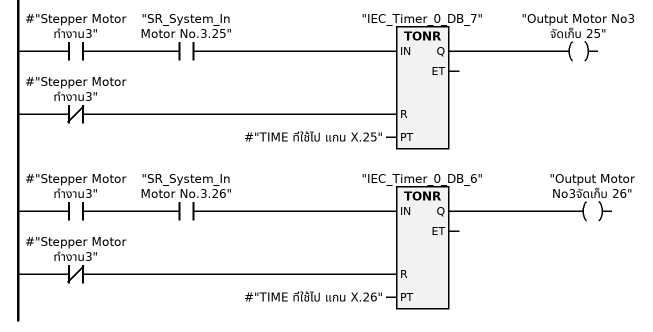
   "IEC_Timer_0_DB_1".TONR(IN := #"Stepper Motor  ทำงาน3" AND "SR_System_In Motor No.3.1",
                           R := NOT #"Stepper Motor  ทำงาน3",
                           PT := #"TIME ที่ใช้ไป แกน X.1");
   "Output Motor No3 จัดเก็บ 1" := "IEC_Timer_0_DB_1".Q;
   "IEC_Timer_0_DB_4".TONR(IN := #"Stepper Motor  ทำงาน3" AND "SR_System_In Motor No.3.2",
                           R := NOT #"Stepper Motor  ทำงาน3",
                           PT := #"TIME ที่ใช้ไป แกน X.2");
   "Output Motor No3 จัดเก็บ 2" := "IEC_Timer_0_DB_4".Q;
   "IEC_Timer_0_DB_5".TONR(IN := #"Stepper Motor  ทำงาน3" AND "SR_System_In Motor No.3.3",
                           R := NOT #"Stepper Motor  ทำงาน3",
                           PT := #"TIME ที่ใช้ไป แกน X.3");
   "Output Motor No3จัดเก็บ 3" := "IEC_Timer_0_DB_5".Q;
   "IEC_Timer_0_DB_28".TONR(IN := #"Stepper Motor  ทำงาน3" AND "SR_System_In Motor No.3.4",
                           R := NOT #"Stepper Motor  ทำงาน3",
                           PT := #"TIME ที่ใช้ไป แกน X.4");
   "Output Motor No3 จัดเก็บ 4" := "IEC_Timer_0_DB_28".Q;
   "IEC_Timer_0_DB_27".TONR(IN := #"Stepper Motor  ทำงาน3" AND "SR_System_In Motor No.3.5",
                           R := NOT #"Stepper Motor  ทำงาน3",
                           PT := #"TIME ที่ใช้ไป แกน X.5");
   "Output Motor No3จัดเก็บ 5" := "IEC_Timer_0_DB_27".Q;
   "IEC_Timer_0_DB_26".TONR(IN := #"Stepper Motor  ทำงาน3" AND "SR_System_In Motor No.3.6",
                           R := NOT #"Stepper Motor  ทำงาน3",
                           PT := #"TIME ที่ใช้ไป แกน X.6");
   "Output Motor No3 จัดเก็บ 6" := "IEC_Timer_0_DB_26".Q;
   "IEC_Timer_0_DB_25".TONR(IN := #"Stepper Motor  ทำงาน3" AND "SR_System_In Motor No.3.7",
                           R := NOT #"Stepper Motor  ทำงาน3",
                           PT := #"TIME ที่ใช้ไป แกน X.7");
   "Output Motor No3 จัดเก็บ 7" := "IEC_Timer_0_DB_25".Q;
   "IEC_Timer_0_DB_24".TONR(IN := #"Stepper Motor  ทำงาน3" AND "SR_System_In Motor No.3.8",
                           R := NOT #"Stepper Motor  ทำงาน3",
                           PT := #"TIME ที่ใช้ไป แกน X.8");
   "Output Motor No3 จัดเก็บ 8" := "IEC_Timer_0_DB_24".Q;
   "IEC_Timer_0_DB_23".TONR(IN := #"Stepper Motor  ทำงาน3" AND "SR_System_In Motor No.3.9",
                           R := NOT #"Stepper Motor  ทำงาน3",
                           PT := #"TIME ที่ใช้ไป แกน X.9");
   "Output Motor No3 จัดเก็บ 9" := "IEC_Timer_0_DB_23".Q;
   "IEC_Timer_0_DB_22".TONR(IN := #"Stepper Motor  ทำงาน3" AND "SR_System_In Motor No.3.10",
                           R := NOT #"Stepper Motor  ทำงาน3",
                           PT := #"TIME ที่ใช้ไป แกน X.10");
   "Output Motor No3 จัดเก็บ10" := "IEC_Timer_0_DB_22".Q;
   "IEC_Timer_0_DB_21".TONR(IN := #"Stepper Motor  ทำงาน3" AND "SR_System_In Motor No.3.11",
                           R := NOT #"Stepper Motor  ทำงาน3",
                           PT := #"TIME ที่ใช้ไป แกน X.11");
   "Output Motor No3จัดเก็บ 11" := "IEC_Timer_0_DB_21".Q;
   "IEC_Timer_0_DB_20".TONR(IN := #"Stepper Motor  ทำงาน3" AND "SR_System_In Motor No.3.12",
                           R := NOT #"Stepper Motor  ทำงาน3",
                           PT := #"TIME ที่ใช้ไป แกน X.12");
   "Output Motor No3 จัดเก็บ 12" := "IEC_Timer_0_DB_20".Q;
   "IEC_Timer_0_DB_19".TONR(IN := #"Stepper Motor  ทำงาน3" AND "SR_System_In Motor No.3.13",
                           R := NOT #"Stepper Motor  ทำงาน3",
                           PT := #"TIME ที่ใช้ไป แกน X.13");
   "Output Motor No3จัดเก็บ 13" := "IEC_Timer_0_DB_19".Q;
   "IEC_Timer_0_DB_18".TONR(IN := #"Stepper Motor  ทำงาน3" AND "SR_System_In Motor No.3.14",
                           R := NOT #"Stepper Motor  ทำงาน3",
                           PT := #"TIME ที่ใช้ไป แกน X.14");
   "Output Motor No3 จัดเก็บ 14" := "IEC_Timer_0_DB_18".Q;
   "IEC_Timer_0_DB_17".TONR(IN := #"Stepper Motor  ทำงาน3" AND "SR_System_In Motor No.3.15",
                           R := NOT #"Stepper Motor  ทำงาน3",
                           PT := #"TIME ที่ใช้ไป แกน X.15");
   "Output Motor No3 จัดเก็บ 15" := "IEC_Timer_0_DB_17".Q;
   "IEC_Timer_0_DB_16".TONR(IN := #"Stepper Motor  ทำงาน3" AND "SR_System_In Motor No.3.16",
                           R := NOT #"Stepper Motor  ทำงาน3",
                           PT := #"TIME ที่ใช้ไป แกน X.16");
   "Output Motor No3 จัดเก็บ 16" := "IEC_Timer_0_DB_16".Q;
   "IEC_Timer_0_DB_15".TONR(IN := #"Stepper Motor  ทำงาน3" AND "SR_System_In Motor No.3.17",
                           R := NOT #"Stepper Motor  ทำงาน3",
                           PT := #"TIME ที่ใช้ไป แกน X.17");
   "Output Motor No3 จัดเก็บ 17" := "IEC_Timer_0_DB_15".Q;
   "IEC_Timer_0_DB_14".TONR(IN := #"Stepper Motor  ทำงาน3" AND "SR_System_In Motor No.3.18",
                           R := NOT #"Stepper Motor  ทำงาน3",
                           PT := #"TIME ที่ใช้ไป แกน X.18");
   "Output Motor No3 จัดเก็บ 18" := "IEC_Timer_0_DB_14".Q;
   "IEC_Timer_0_DB_13".TONR(IN := #"Stepper Motor  ทำงาน3" AND "SR_System_In Motor No.3.19",
                           R := NOT #"Stepper Motor  ทำงาน3",
                           PT := #"TIME ที่ใช้ไป แกน X.19");
   "Output Motor No3จัดเก็บ 19" := "IEC_Timer_0_DB_13".Q;
   "IEC_Timer_0_DB_12".TONR(IN := #"Stepper Motor  ทำงาน3" AND "SR_System_In Motor No.3.20",
                           R := NOT #"Stepper Motor  ทำงาน3",
                           PT := #"TIME ที่ใช้ไป แกน X.20");
   "Output Motor No3 จัดเก็บ 20" := "IEC_Timer_0_DB_12".Q;
   "IEC_Timer_0_DB_11".TONR(IN := #"Stepper Motor  ทำงาน3" AND "SR_System_In Motor No.3.21",
                           R := NOT #"Stepper Motor  ทำงาน3",
                           PT := #"TIME ที่ใช้ไป แกน X.21");
   "Output Motor No3จัดเก็บ 21" := "IEC_Timer_0_DB_11".Q;
   "IEC_Timer_0_DB_10".TONR(IN := #"Stepper Motor  ทำงาน3" AND "SR_System_In Motor No.3.22",
                           R := NOT #"Stepper Motor  ทำงาน3",
                           PT := #"TIME ที่ใช้ไป แกน X.22");
   "Output Motor No3 จัดเก็บ 22" := "IEC_Timer_0_DB_10".Q;
   "IEC_Timer_0_DB_9".TONR(IN := #"Stepper Motor  ทำงาน3" AND "SR_System_In Motor No.3.23",
                           R := NOT #"Stepper Motor  ทำงาน3",
                           PT := #"TIME ที่ใช้ไป แกน X.23");
   "Output Motor No3 จัดเก็บ 23" := "IEC_Timer_0_DB_9".Q;
   "IEC_Timer_0_DB_8".TONR(IN := #"Stepper Motor  ทำงาน3" AND "SR_System_In Motor No.3.24",
                           R := NOT #"Stepper Motor  ทำงาน3",
                           PT := #"TIME ที่ใช้ไป แกน X.24");
   "Output Motor No3จัดเก็บ 24" := "IEC_Timer_0_DB_8".Q;
   "IEC_Timer_0_DB_7".TONR(IN := #"Stepper Motor  ทำงาน3" AND "SR_System_In Motor No.3.25",
                           R := NOT #"Stepper Motor  ทำงาน3",
                           PT := #"TIME ที่ใช้ไป แกน X.25");
   "Output Motor No3 จัดเก็บ 25" := "IEC_Timer_0_DB_7".Q;
   "IEC_Timer_0_DB_6".TONR(IN := #"Stepper Motor  ทำงาน3" AND "SR_System_In Motor No.3.26",
                           R := NOT #"Stepper Motor  ทำงาน3",
                           PT := #"TIME ที่ใช้ไป แกน X.26");
   "Output Motor No3จัดเก็บ 26" := "IEC_Timer_0_DB_6".Q;
END_REGION

REGION Network 3
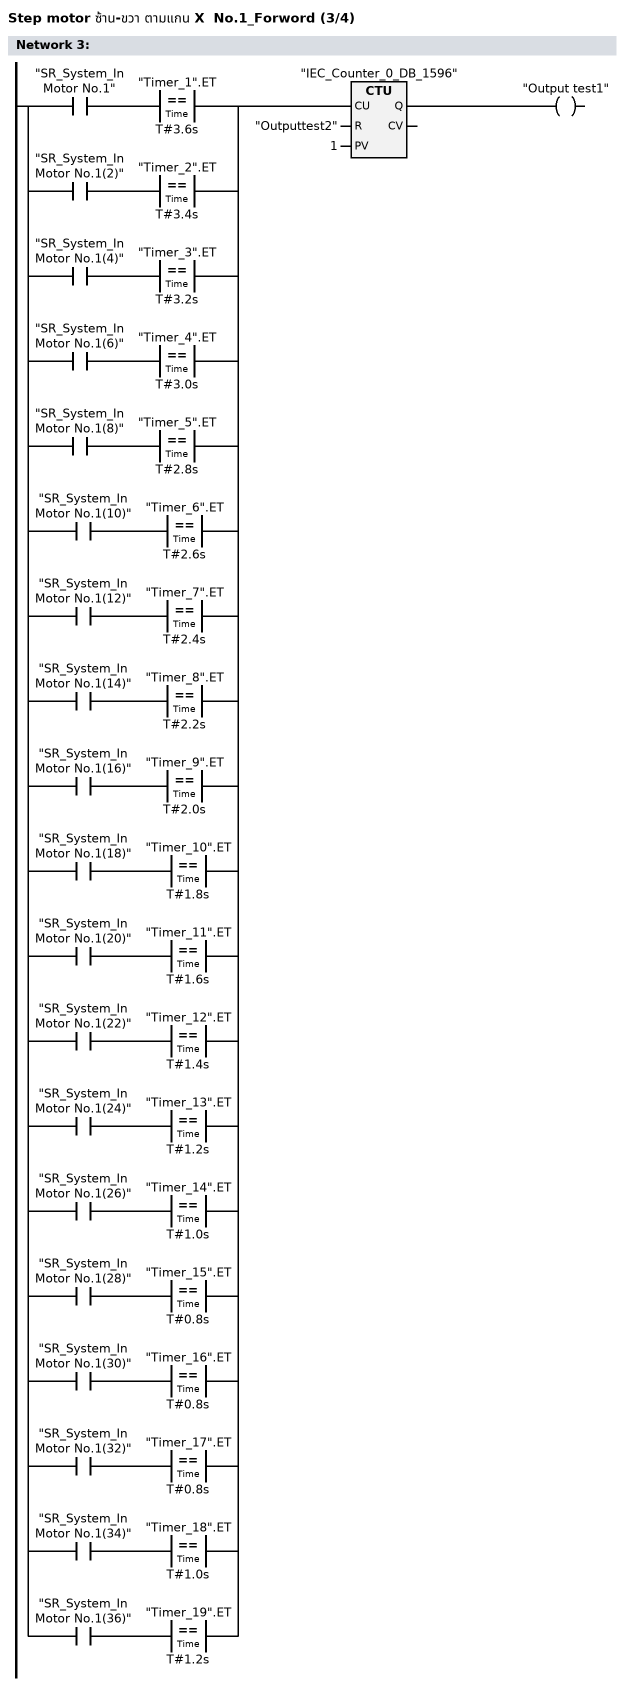
   "IEC_Counter_0_DB_1596".CTU(CU := ("SR_System_In Motor No.1" AND ("Timer_1".ET = T#3.6s)) OR ("SR_System_In Motor No.1(2)" AND ("Timer_2".ET = T#3.4s)) OR ("SR_System_In Motor No.1(4)" AND ("Timer_3".ET = T#3.2s)) OR ("SR_System_In Motor No.1(6)" AND ("Timer_4".ET = T#3.0s)) OR ("SR_System_In Motor No.1(8)" AND ("Timer_5".ET = T#2.8s)) OR ("SR_System_In Motor No.1(10)" AND ("Timer_6".ET = T#2.6s)) OR ("SR_System_In Motor No.1(12)" AND ("Timer_7".ET = T#2.4s)) OR ("SR_System_In Motor No.1(14)" AND ("Timer_8".ET = T#2.2s)) OR ("SR_System_In Motor No.1(16)" AND ("Timer_9".ET = T#2.0s)) OR ("SR_System_In Motor No.1(18)" AND ("Timer_10".ET = T#1.8s)) OR ("SR_System_In Motor No.1(20)" AND ("Timer_11".ET = T#1.6s)) OR ("SR_System_In Motor No.1(22)" AND ("Timer_12".ET = T#1.4s)) OR ("SR_System_In Motor No.1(24)" AND ("Timer_13".ET = T#1.2s)) OR ("SR_System_In Motor No.1(26)" AND ("Timer_14".ET = T#1.0s)) OR ("SR_System_In Motor No.1(28)" AND ("Timer_15".ET = T#0.8s)) OR ("SR_System_In Motor No.1(30)" AND ("Timer_16".ET = T#0.8s)) OR ("SR_System_In Motor No.1(32)" AND ("Timer_17".ET = T#0.8s)) OR ("SR_System_In Motor No.1(34)" AND ("Timer_18".ET = T#1.0s)) OR ("SR_System_In Motor No.1(36)" AND ("Timer_19".ET = T#1.2s)),
                           R := "Outputtest2",
                           PV := 1);
   "Output test1" := "IEC_Counter_0_DB_1596".Q;
END_REGION

REGION Network 4
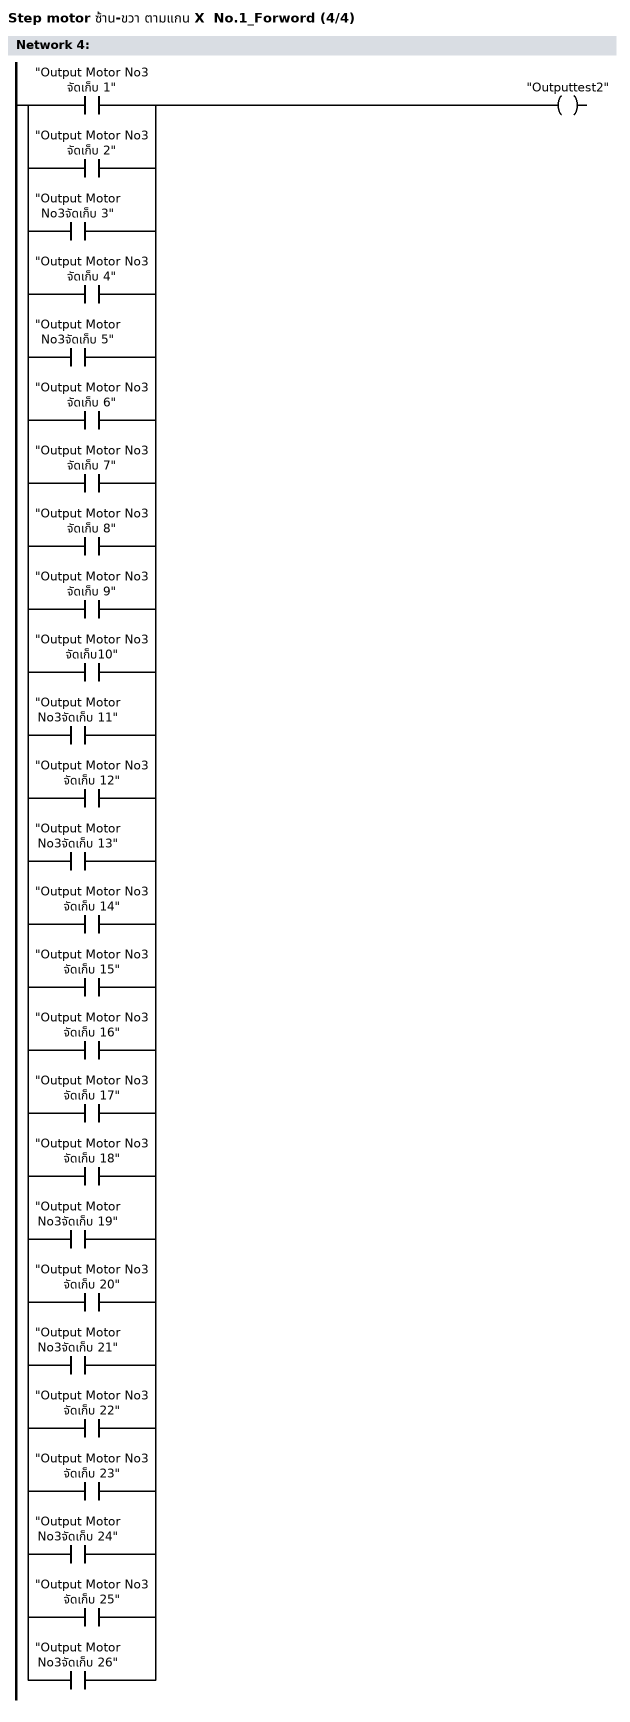
   RUNG wire#powerrail
      Contact( "Output Motor No3 จัดเก็บ 1" )
      wire#w1
      Coil( "Outputtest2" )
   END_RUNG
   RUNG wire#powerrail
      Contact( "Output Motor No3 จัดเก็บ 2" )
   END_RUNG wire#w1
   RUNG wire#powerrail
      Contact( "Output Motor No3จัดเก็บ 3" )
   END_RUNG wire#w1
   RUNG wire#powerrail
      Contact( "Output Motor No3 จัดเก็บ 4" )
   END_RUNG wire#w1
   RUNG wire#powerrail
      Contact( "Output Motor No3จัดเก็บ 5" )
   END_RUNG wire#w1
   RUNG wire#powerrail
      Contact( "Output Motor No3 จัดเก็บ 6" )
   END_RUNG wire#w1
   RUNG wire#powerrail
      Contact( "Output Motor No3 จัดเก็บ 7" )
   END_RUNG wire#w1
   RUNG wire#powerrail
      Contact( "Output Motor No3 จัดเก็บ 8" )
   END_RUNG wire#w1
   RUNG wire#powerrail
      Contact( "Output Motor No3 จัดเก็บ 9" )
   END_RUNG wire#w1
   RUNG wire#powerrail
      Contact( "Output Motor No3 จัดเก็บ10" )
   END_RUNG wire#w1
   RUNG wire#powerrail
      Contact( "Output Motor No3จัดเก็บ 11" )
   END_RUNG wire#w1
   RUNG wire#powerrail
      Contact( "Output Motor No3 จัดเก็บ 12" )
   END_RUNG wire#w1
   RUNG wire#powerrail
      Contact( "Output Motor No3จัดเก็บ 13" )
   END_RUNG wire#w1
   RUNG wire#powerrail
      Contact( "Output Motor No3 จัดเก็บ 14" )
   END_RUNG wire#w1
   RUNG wire#powerrail
      Contact( "Output Motor No3 จัดเก็บ 15" )
   END_RUNG wire#w1
   RUNG wire#powerrail
      Contact( "Output Motor No3 จัดเก็บ 16" )
   END_RUNG wire#w1
   RUNG wire#powerrail
      Contact( "Output Motor No3 จัดเก็บ 17" )
   END_RUNG wire#w1
   RUNG wire#powerrail
      Contact( "Output Motor No3 จัดเก็บ 18" )
   END_RUNG wire#w1
   RUNG wire#powerrail
      Contact( "Output Motor No3จัดเก็บ 19" )
   END_RUNG wire#w1
   RUNG wire#powerrail
      Contact( "Output Motor No3 จัดเก็บ 20" )
   END_RUNG wire#w1
   RUNG wire#powerrail
      Contact( "Output Motor No3จัดเก็บ 21" )
   END_RUNG wire#w1
   RUNG wire#powerrail
      Contact( "Output Motor No3 จัดเก็บ 22" )
   END_RUNG wire#w1
   RUNG wire#powerrail
      Contact( "Output Motor No3 จัดเก็บ 23" )
   END_RUNG wire#w1
   RUNG wire#powerrail
      Contact( "Output Motor No3จัดเก็บ 24" )
   END_RUNG wire#w1
   RUNG wire#powerrail
      Contact( "Output Motor No3 จัดเก็บ 25" )
   END_RUNG wire#w1
   RUNG wire#powerrail
      Contact( "Output Motor No3จัดเก็บ 26" )
   END_RUNG wire#w1
   // the same network as SCL:
   "Outputtest2" := "Output Motor No3 จัดเก็บ 1" OR "Output Motor No3 จัดเก็บ 2" OR "Output Motor No3จัดเก็บ 3" OR "Output Motor No3 จัดเก็บ 4" OR "Output Motor No3จัดเก็บ 5" OR "Output Motor No3 จัดเก็บ 6" OR "Output Motor No3 จัดเก็บ 7" OR "Output Motor No3 จัดเก็บ 8" OR "Output Motor No3 จัดเก็บ 9" OR "Output Motor No3 จัดเก็บ10" OR "Output Motor No3จัดเก็บ 11" OR "Output Motor No3 จัดเก็บ 12" OR "Output Motor No3จัดเก็บ 13" OR "Output Motor No3 จัดเก็บ 14" OR "Output Motor No3 จัดเก็บ 15" OR "Output Motor No3 จัดเก็บ 16" OR "Output Motor No3 จัดเก็บ 17" OR "Output Motor No3 จัดเก็บ 18" OR "Output Motor No3จัดเก็บ 19" OR "Output Motor No3 จัดเก็บ 20" OR "Output Motor No3จัดเก็บ 21" OR "Output Motor No3 จัดเก็บ 22" OR "Output Motor No3 จัดเก็บ 23" OR "Output Motor No3จัดเก็บ 24" OR "Output Motor No3 จัดเก็บ 25" OR "Output Motor No3จัดเก็บ 26";
END_REGION
END_FUNCTION_BLOCK

FUNCTION_BLOCK "Step motor ซ้าย-ขวา ตามแกน X No.1_Blackword"   // FB6, LAD
{ S7_Optimized_Access := 'TRUE' }
VERSION : 0.1
   VAR_INPUT
      "TIME ที่ใช้ จาก แกน X.1 ไปจุดเริ่มต้น" : Time;
      "TIME ที่ใช้ จาก แกน X.2 ไปจุดเริ่มต้น" : Time;
      "TIME ที่ใช้ จาก แกน X.3 ไปจุดเริ่มต้น" : Time;
      "TIME ที่ใช้ จาก แกน X.4 ไปจุดเริ่มต้น" : Time;
      "TIME ที่ใช้ จาก แกน X.5 ไปจุดเริ่มต้น" : Time;
      "TIME ที่ใช้ จาก แกน X.6 ไปจุดเริ่มต้น" : Time;
      "TIME ที่ใช้ จาก แกน X.7 ไปจุดเริ่มต้น" : Time;
      "TIME ที่ใช้ จาก แกน X.8 ไปจุดเริ่มต้น" : Time;
      "TIME ที่ใช้ จาก แกน X.9 ไปจุดเริ่มต้น" : Time;
      "TIME ที่ใช้ จาก แกน X.10 ไปจุดเริ่มต้น" : Time;
      "TIME ที่ใช้ จาก แกน X.11 ไปจุดเริ่มต้น" : Time;
      "TIME ที่ใช้ จาก แกน X.12 ไปจุดเริ่มต้น" : Time;
      "TIME ที่ใช้ จาก แกน X.13 ไปจุดเริ่มต้น" : Time;
      "TIME ที่ใช้ จาก แกน X.14 ไปจุดเริ่มต้น" : Time;
      "TIME ที่ใช้ จาก แกน X.15 ไปจุดเริ่มต้น" : Time;
      "TIME ที่ใช้ จาก แกน X.16 ไปจุดเริ่มต้น" : Time;
      "TIME ที่ใช้ จาก แกน X.17 ไปจุดเริ่มต้น" : Time;
      "TIME ที่ใช้ จาก แกน X.18 ไปจุดเริ่มต้น" : Time;
      "TIME ที่ใช้ จาก แกน X.19 ไปจุดเริ่มต้น" : Time;
      "TIME ที่ใช้ จาก แกน X.20 ไปจุดเริ่มต้น" : Time;
      "TIME ที่ใช้ จาก แกน X.21 ไปจุดเริ่มต้น" : Time;
      "TIME ที่ใช้ จาก แกน X.22 ไปจุดเริ่มต้น" : Time;
      "TIME ที่ใช้ จาก แกน X.23 ไปจุดเริ่มต้น" : Time;
      "TIME ที่ใช้ จาก แกน X.24 ไปจุดเริ่มต้น" : Time;
      "TIME ที่ใช้ จาก แกน X.25 ไปจุดเริ่มต้น" : Time;
      "TIME ที่ใช้ จาก แกน X.26 ไปจุดเริ่มต้น" : Time;
   END_VAR
   VAR_IN_OUT
      "Step motor  Backword ทำงาน No.3" : Bool;
   END_VAR
   VAR_TEMP   // added for the SCL form of the ladder/FBD networks
      _w1 : Bool;
      _w2 : Bool;
      _w3 : Bool;
      _w4 : Bool;
      _w5 : Bool;
      _w6 : Bool;
      _w7 : Bool;
      _w8 : Bool;
      _w9 : Bool;
      _w10 : Bool;
      _w11 : Bool;
      _w12 : Bool;
      _w13 : Bool;
      _w14 : Bool;
      _w15 : Bool;
      _w16 : Bool;
      _w17 : Bool;
      _w18 : Bool;
      _w19 : Bool;
      _w20 : Bool;
      _w21 : Bool;
      _w22 : Bool;
      _w23 : Bool;
      _w24 : Bool;
      _w25 : Bool;
      _w26 : Bool;
      _w27 : Bool;
      _w28 : Bool;
      _w29 : Bool;
      _w30 : Bool;
      _w31 : Bool;
      _w32 : Bool;
      _w33 : Bool;
      _w34 : Bool;
      _w35 : Bool;
      _w36 : Bool;
      _w37 : Bool;
      _w38 : Bool;
      _w39 : Bool;
      _w40 : Bool;
      _w41 : Bool;
      _w42 : Bool;
      _w43 : Bool;
      _w44 : Bool;
      _w45 : Bool;
      _w46 : Bool;
      _w47 : Bool;
      _w48 : Bool;
      _w49 : Bool;
      _w50 : Bool;
      _w51 : Bool;
   END_VAR
BEGIN

REGION Network 1
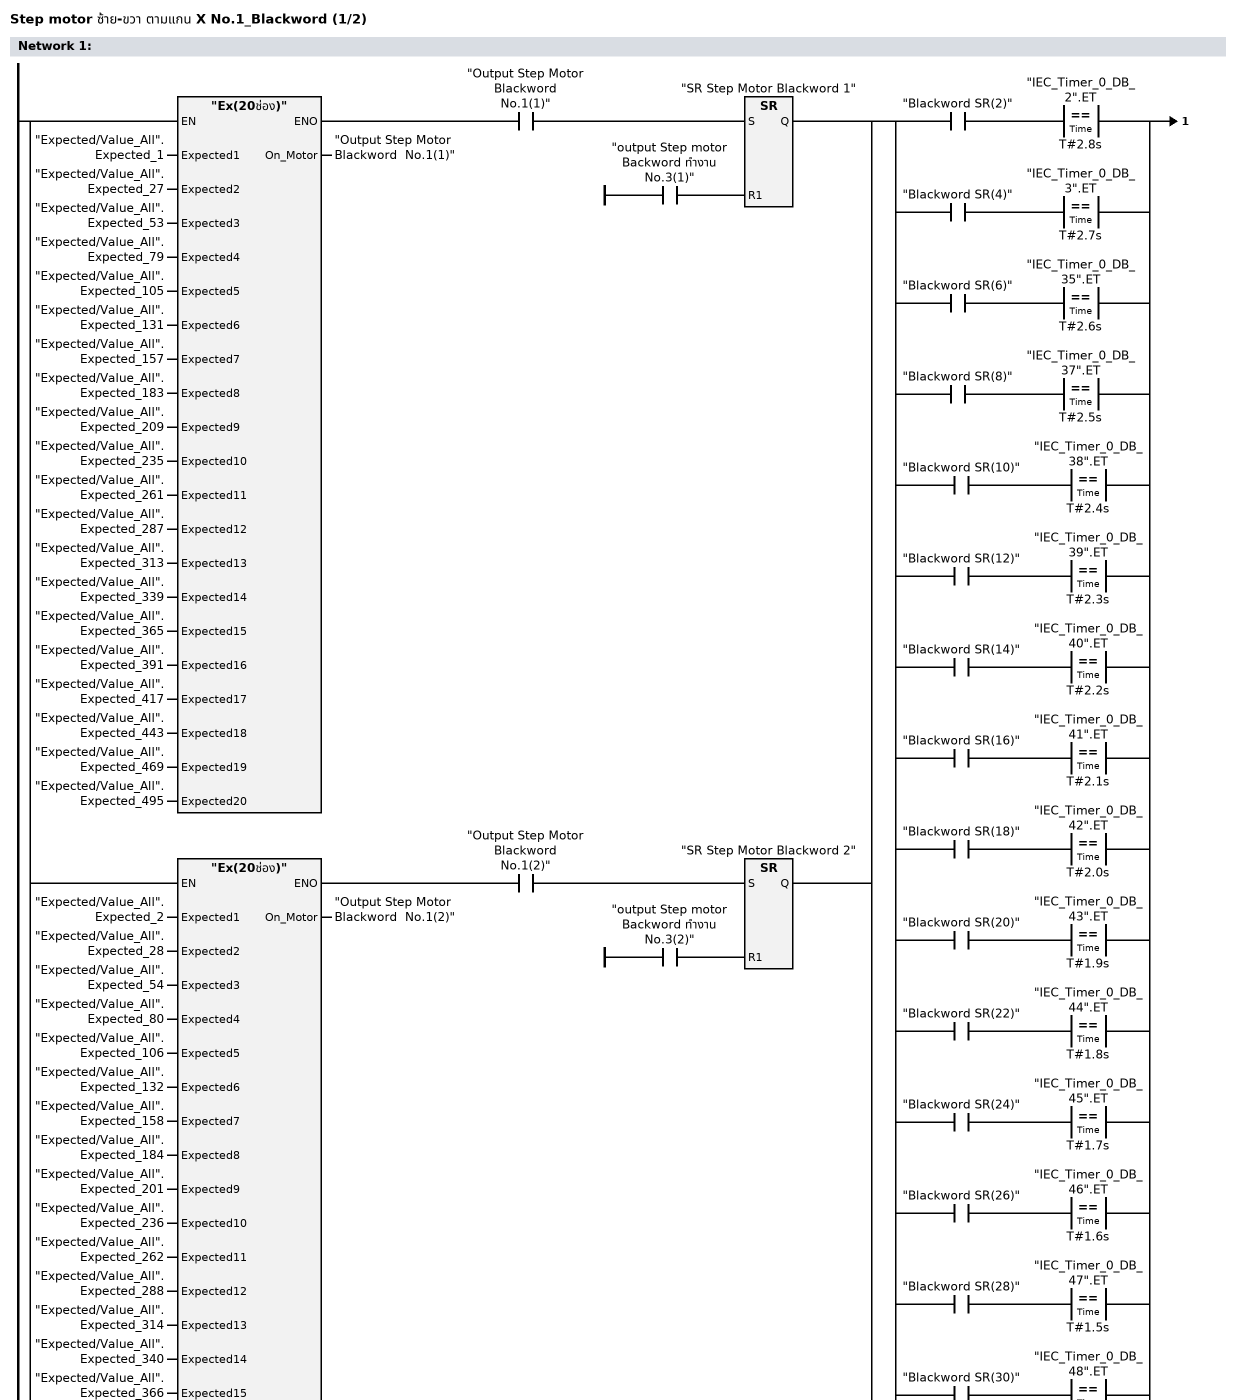
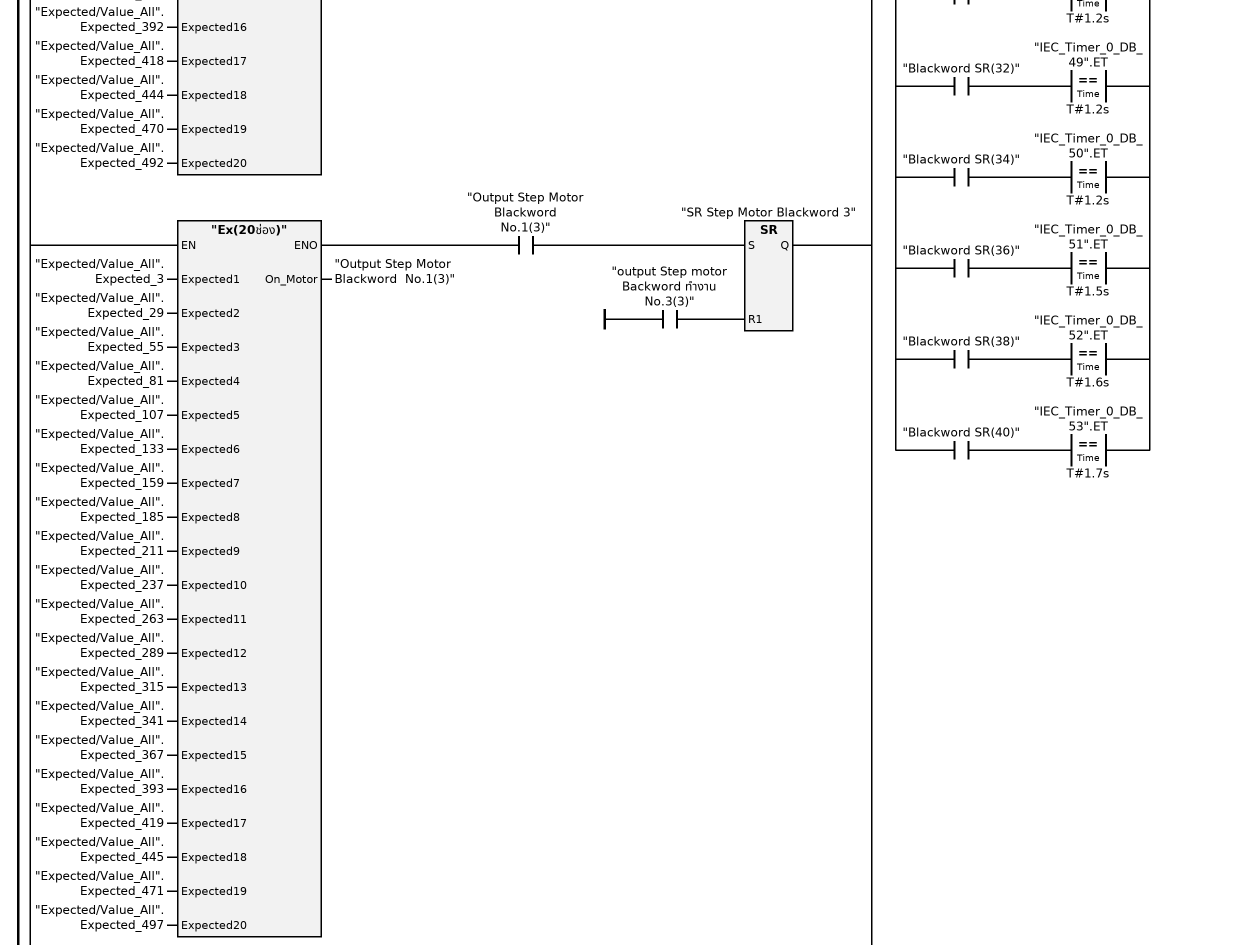
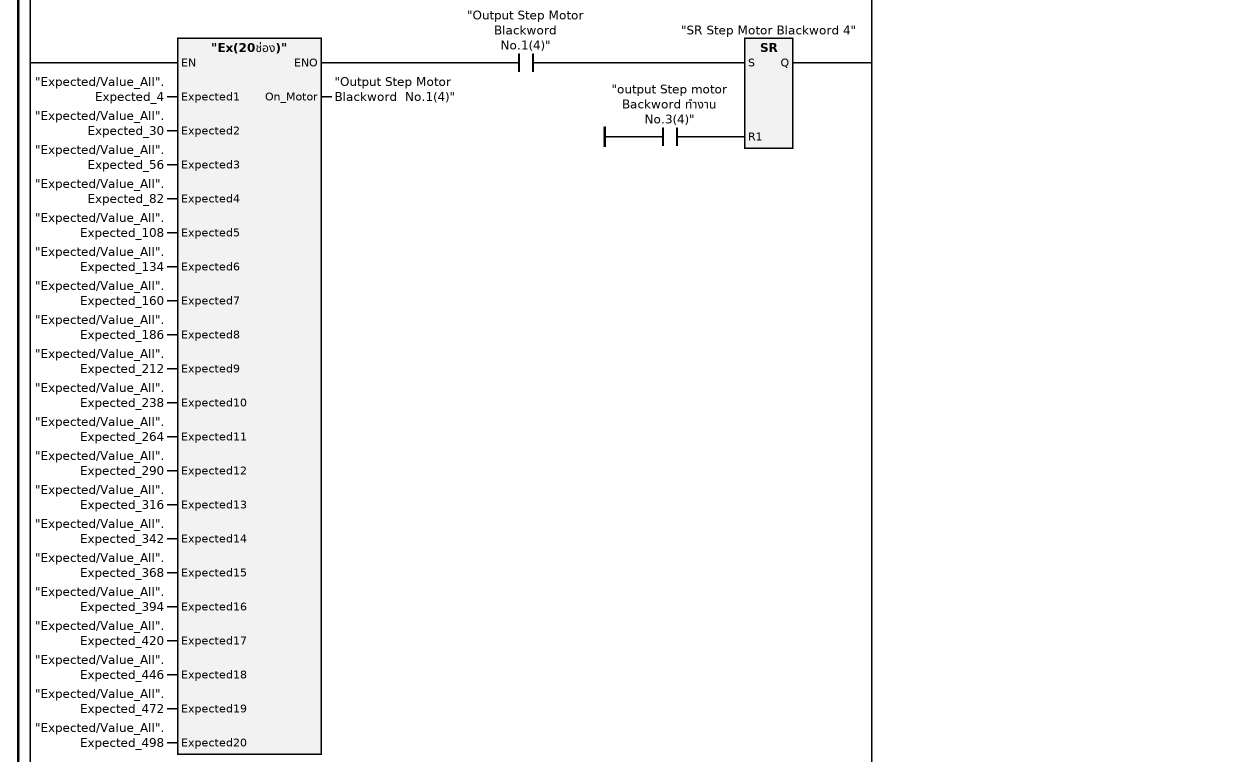
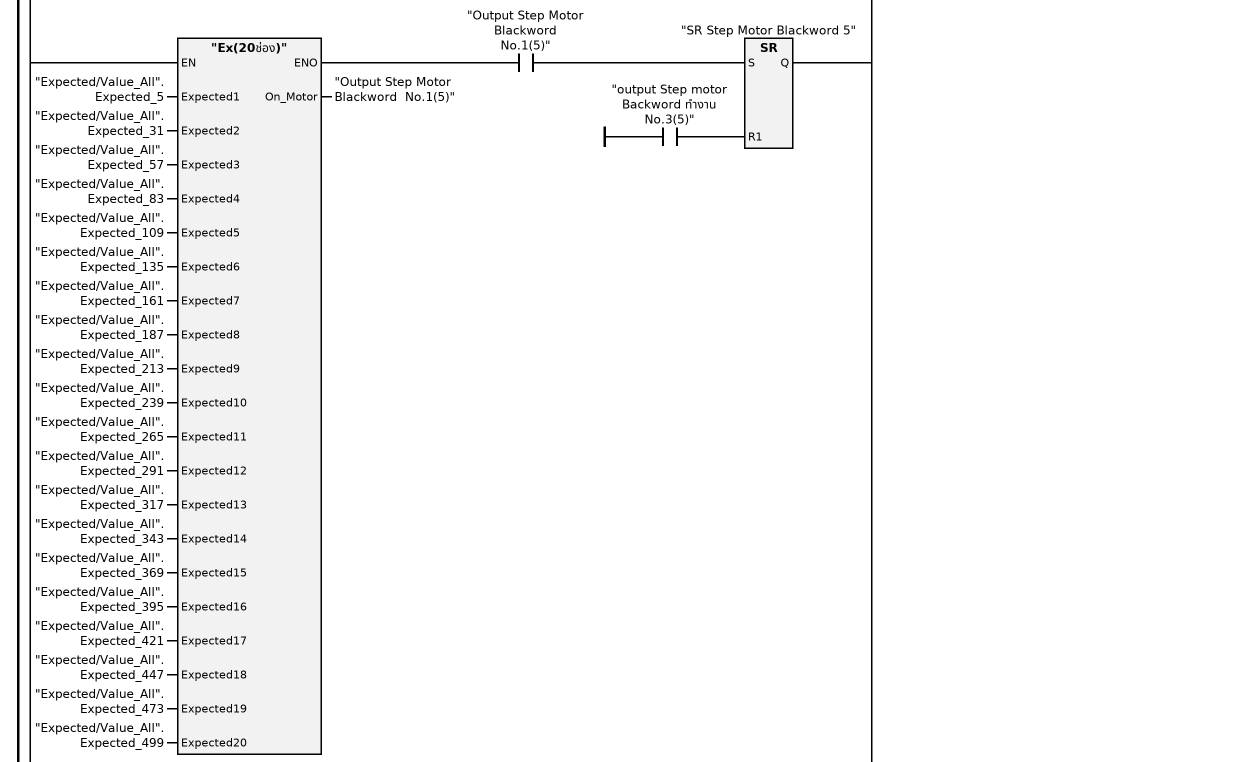
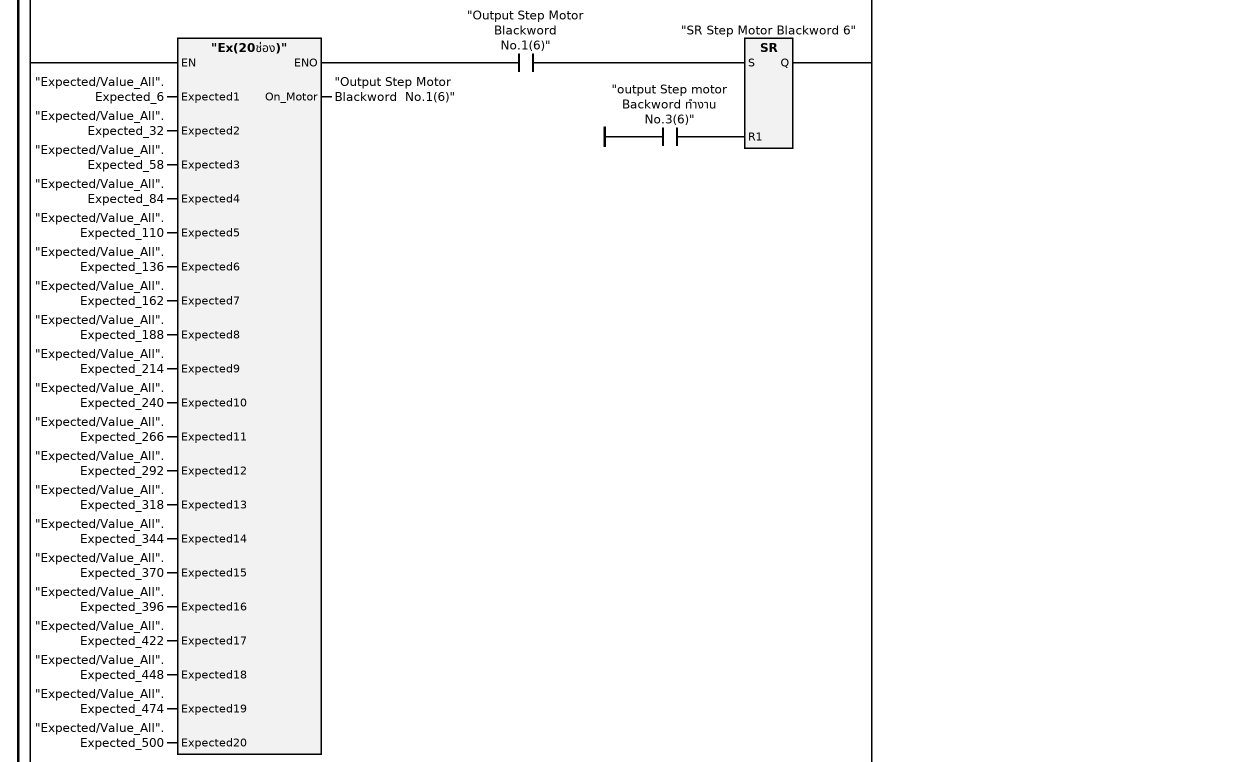
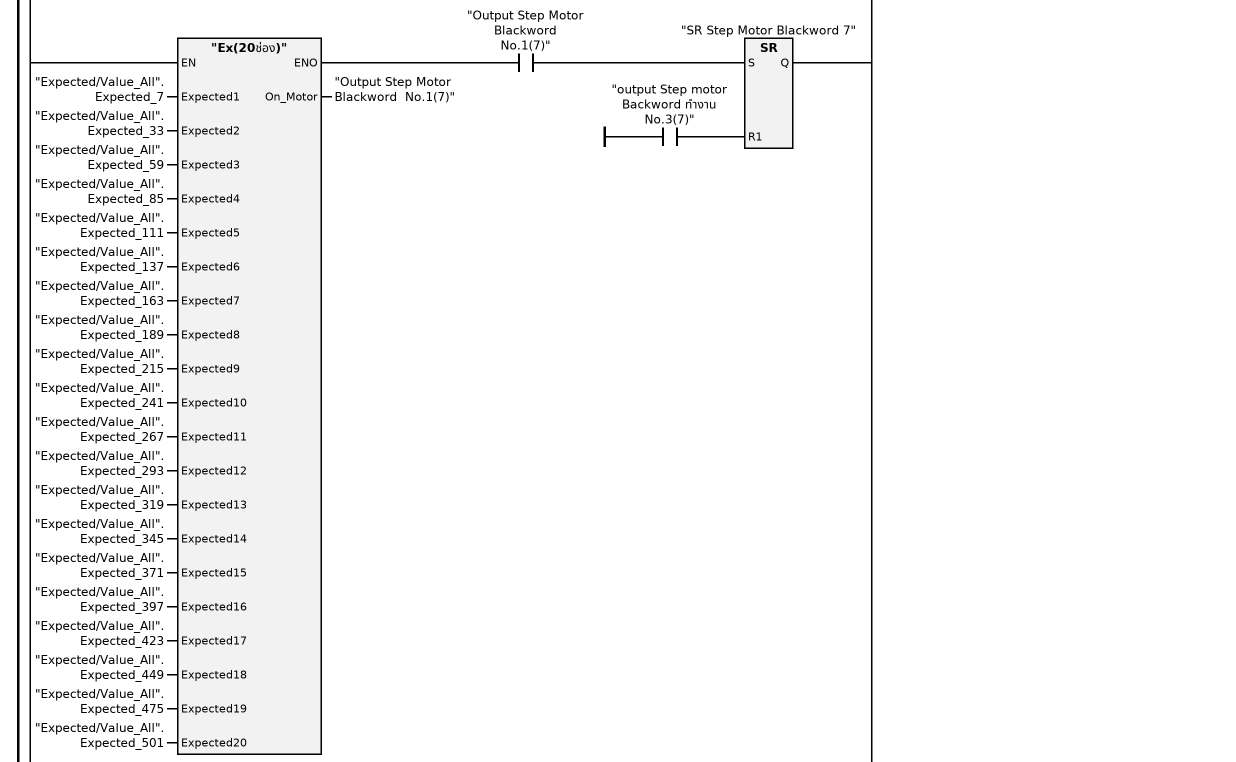
